(* PLC project DsmEasyConfig *)
(* stored: creationDateTime 2022-10-05T09:23:09.683, modificationDateTime 2022-10-05T09:23:09.683 *)

TYPE DFC_rbr_outA01OL : STRUCT
  DTC : UDINT := 16#140100;
  DFCid : UINT := 471;
  debounceMethod : USINT := TIME_UP_DOWN;
END_STRUCT;
END_TYPE

TYPE DFC_rbr_outA01OT : STRUCT
  DTC : UDINT := 16#140200;
  DFCid : UINT := 472;
  debounceMethod : USINT := TIME_UP_DOWN;
END_STRUCT;
END_TYPE

TYPE DFC_rbr_outA01SCB : STRUCT
  DTC : UDINT := 16#140300;
  DFCid : UINT := 473;
  debounceMethod : USINT := TIME_UP_DOWN;
END_STRUCT;
END_TYPE

TYPE DFC_rbr_outA02OC : STRUCT
  DTC : UDINT := 16#140500;
  DFCid : UINT := 971;
  debounceMethod : USINT := NO_DEBOUNCE;
END_STRUCT;
END_TYPE

TYPE DFC_rbr_outA01SCG : STRUCT
  DTC : UDINT := 16#140400;
  DFCid : UINT := 474;
  debounceMethod : USINT := TIME_UP_DOWN;
END_STRUCT;
END_TYPE

TYPE DFC_rbr_outA02OL : STRUCT
  DTC : UDINT := 16#140600;
  DFCid : UINT := 475;
  debounceMethod : USINT := TIME_UP_DOWN;
END_STRUCT;
END_TYPE

TYPE DFC_rbr_outA02OR : STRUCT
  DTC : UDINT := 16#140700;
  DFCid : UINT := 476;
  debounceMethod : USINT := TIME_UP_DOWN;
END_STRUCT;
END_TYPE

TYPE DFC_rbr_outA02OT : STRUCT
  DTC : UDINT := 16#140800;
  DFCid : UINT := 477;
  debounceMethod : USINT := TIME_UP_DOWN;
END_STRUCT;
END_TYPE

TYPE DFC_rbr_outA02SCB : STRUCT
  DTC : UDINT := 16#140900;
  DFCid : UINT := 478;
  debounceMethod : USINT := TIME_UP_DOWN;
END_STRUCT;
END_TYPE

TYPE DFC_rbr_outA02SCG : STRUCT
  DTC : UDINT := 16#140A00;
  DFCid : UINT := 479;
  debounceMethod : USINT := TIME_UP_DOWN;
END_STRUCT;
END_TYPE

TYPE DFC_rbr_outA03OC : STRUCT
  DTC : UDINT := 16#140B00;
  DFCid : UINT := 973;
  debounceMethod : USINT := NO_DEBOUNCE;
END_STRUCT;
END_TYPE

TYPE DFC_rbr_outA03OL : STRUCT
  DTC : UDINT := 16#140C00;
  DFCid : UINT := 480;
  debounceMethod : USINT := TIME_UP_DOWN;
END_STRUCT;
END_TYPE

TYPE DFC_rbr_outA03OT : STRUCT
  DTC : UDINT := 16#140D00;
  DFCid : UINT := 481;
  debounceMethod : USINT := TIME_UP_DOWN;
END_STRUCT;
END_TYPE

TYPE DFC_rbr_outA03SCB : STRUCT
  DTC : UDINT := 16#140E00;
  DFCid : UINT := 482;
  debounceMethod : USINT := TIME_UP_DOWN;
END_STRUCT;
END_TYPE

TYPE DFC_rbr_outA03SCG : STRUCT
  DTC : UDINT := 16#140F00;
  DFCid : UINT := 483;
  debounceMethod : USINT := TIME_UP_DOWN;
END_STRUCT;
END_TYPE

TYPE DFC_rbr_outA04OC : STRUCT
  DTC : UDINT := 16#141000;
  DFCid : UINT := 975;
  debounceMethod : USINT := NO_DEBOUNCE;
END_STRUCT;
END_TYPE

TYPE DFC_rbr_outA04OL : STRUCT
  DTC : UDINT := 16#141100;
  DFCid : UINT := 484;
  debounceMethod : USINT := TIME_UP_DOWN;
END_STRUCT;
END_TYPE

TYPE DFC_rbr_outA04OT : STRUCT
  DTC : UDINT := 16#141200;
  DFCid : UINT := 485;
  debounceMethod : USINT := TIME_UP_DOWN;
END_STRUCT;
END_TYPE

TYPE DFC_rbr_outA04SCB : STRUCT
  DTC : UDINT := 16#141300;
  DFCid : UINT := 486;
  debounceMethod : USINT := TIME_UP_DOWN;
END_STRUCT;
END_TYPE

TYPE DFC_rbr_outA04SCG : STRUCT
  DTC : UDINT := 16#141400;
  DFCid : UINT := 487;
  debounceMethod : USINT := TIME_UP_DOWN;
END_STRUCT;
END_TYPE

TYPE DFC_rbr_outA05OC : STRUCT
  DTC : UDINT := 16#141500;
  DFCid : UINT := 977;
  debounceMethod : USINT := NO_DEBOUNCE;
END_STRUCT;
END_TYPE

TYPE DFC_rbr_outA05OL : STRUCT
  DTC : UDINT := 16#141600;
  DFCid : UINT := 488;
  debounceMethod : USINT := TIME_UP_DOWN;
END_STRUCT;
END_TYPE

TYPE DFC_rbr_outA05OR : STRUCT
  DTC : UDINT := 16#141700;
  DFCid : UINT := 489;
  debounceMethod : USINT := TIME_UP_DOWN;
END_STRUCT;
END_TYPE

TYPE DFC_rbr_outA05OT : STRUCT
  DTC : UDINT := 16#141800;
  DFCid : UINT := 490;
  debounceMethod : USINT := TIME_UP_DOWN;
END_STRUCT;
END_TYPE

TYPE DFC_rbr_outA05SCB : STRUCT
  DTC : UDINT := 16#141900;
  DFCid : UINT := 491;
  debounceMethod : USINT := TIME_UP_DOWN;
END_STRUCT;
END_TYPE

TYPE DFC_rbr_outA05SCG : STRUCT
  DTC : UDINT := 16#141A00;
  DFCid : UINT := 492;
  debounceMethod : USINT := TIME_UP_DOWN;
END_STRUCT;
END_TYPE

TYPE DFC_rbr_outA06OR : STRUCT
  DTC : UDINT := 16#141C00;
  DFCid : UINT := 494;
  debounceMethod : USINT := TIME_UP_DOWN;
END_STRUCT;
END_TYPE

TYPE DFC_rbr_outA06OT : STRUCT
  DTC : UDINT := 16#141D00;
  DFCid : UINT := 495;
  debounceMethod : USINT := TIME_UP_DOWN;
END_STRUCT;
END_TYPE

TYPE DFC_rbr_outA06SCB : STRUCT
  DTC : UDINT := 16#141E00;
  DFCid : UINT := 496;
  debounceMethod : USINT := TIME_UP_DOWN;
END_STRUCT;
END_TYPE

TYPE DFC_rbr_outA06SCG : STRUCT
  DTC : UDINT := 16#141F00;
  DFCid : UINT := 497;
  debounceMethod : USINT := TIME_UP_DOWN;
END_STRUCT;
END_TYPE

TYPE DFC_rbr_outA07OC : STRUCT
  DTC : UDINT := 16#142000;
  DFCid : UINT := 979;
  debounceMethod : USINT := NO_DEBOUNCE;
END_STRUCT;
END_TYPE

TYPE DFC_rbr_outA07OL : STRUCT
  DTC : UDINT := 16#142100;
  DFCid : UINT := 498;
  debounceMethod : USINT := TIME_UP_DOWN;
END_STRUCT;
END_TYPE

TYPE DFC_rbr_outA07OT : STRUCT
  DTC : UDINT := 16#142200;
  DFCid : UINT := 499;
  debounceMethod : USINT := TIME_UP_DOWN;
END_STRUCT;
END_TYPE

TYPE DFC_rbr_outA07SCB : STRUCT
  DTC : UDINT := 16#142300;
  DFCid : UINT := 500;
  debounceMethod : USINT := TIME_UP_DOWN;
END_STRUCT;
END_TYPE

TYPE DFC_rbr_outA07SCG : STRUCT
  DTC : UDINT := 16#142400;
  DFCid : UINT := 501;
  debounceMethod : USINT := TIME_UP_DOWN;
END_STRUCT;
END_TYPE

TYPE DFC_rbr_outA08OC : STRUCT
  DTC : UDINT := 16#142500;
  DFCid : UINT := 981;
  debounceMethod : USINT := NO_DEBOUNCE;
END_STRUCT;
END_TYPE

TYPE DFC_rbr_outA08OL : STRUCT
  DTC : UDINT := 16#142600;
  DFCid : UINT := 502;
  debounceMethod : USINT := TIME_UP_DOWN;
END_STRUCT;
END_TYPE

TYPE DFC_rbr_outA08OT : STRUCT
  DTC : UDINT := 16#142700;
  DFCid : UINT := 503;
  debounceMethod : USINT := TIME_UP_DOWN;
END_STRUCT;
END_TYPE

TYPE DFC_rbr_outA08SCB : STRUCT
  DTC : UDINT := 16#142800;
  DFCid : UINT := 504;
  debounceMethod : USINT := TIME_UP_DOWN;
END_STRUCT;
END_TYPE

TYPE DFC_rbr_outA08SCG : STRUCT
  DTC : UDINT := 16#142900;
  DFCid : UINT := 505;
  debounceMethod : USINT := TIME_UP_DOWN;
END_STRUCT;
END_TYPE

TYPE DFC_rbr_outA09OC : STRUCT
  DTC : UDINT := 16#142A00;
  DFCid : UINT := 983;
  debounceMethod : USINT := NO_DEBOUNCE;
END_STRUCT;
END_TYPE

TYPE DFC_rbr_outA09OL : STRUCT
  DTC : UDINT := 16#142B00;
  DFCid : UINT := 506;
  debounceMethod : USINT := TIME_UP_DOWN;
END_STRUCT;
END_TYPE

TYPE DFC_rbr_outA09OR : STRUCT
  DTC : UDINT := 16#142C00;
  DFCid : UINT := 507;
  debounceMethod : USINT := TIME_UP_DOWN;
END_STRUCT;
END_TYPE

TYPE DFC_rbr_outA09OT : STRUCT
  DTC : UDINT := 16#142D00;
  DFCid : UINT := 508;
  debounceMethod : USINT := TIME_UP_DOWN;
END_STRUCT;
END_TYPE

TYPE DFC_rbr_outA09SCB : STRUCT
  DTC : UDINT := 16#142E00;
  DFCid : UINT := 509;
  debounceMethod : USINT := TIME_UP_DOWN;
END_STRUCT;
END_TYPE

TYPE DFC_rbr_outA09SCG : STRUCT
  DTC : UDINT := 16#142F00;
  DFCid : UINT := 510;
  debounceMethod : USINT := TIME_UP_DOWN;
END_STRUCT;
END_TYPE

TYPE DFC_rbr_outA10OC : STRUCT
  DTC : UDINT := 16#143000;
  DFCid : UINT := 985;
  debounceMethod : USINT := NO_DEBOUNCE;
END_STRUCT;
END_TYPE

TYPE DFC_rbr_outA10OL : STRUCT
  DTC : UDINT := 16#143100;
  DFCid : UINT := 511;
  debounceMethod : USINT := TIME_UP_DOWN;
END_STRUCT;
END_TYPE

TYPE DFC_rbr_outA10OT : STRUCT
  DTC : UDINT := 16#143200;
  DFCid : UINT := 512;
  debounceMethod : USINT := TIME_UP_DOWN;
END_STRUCT;
END_TYPE

TYPE DFC_rbr_outA10SCB : STRUCT
  DTC : UDINT := 16#143300;
  DFCid : UINT := 513;
  debounceMethod : USINT := TIME_UP_DOWN;
END_STRUCT;
END_TYPE

TYPE DFC_rbr_outA10SCG : STRUCT
  DTC : UDINT := 16#143400;
  DFCid : UINT := 514;
  debounceMethod : USINT := TIME_UP_DOWN;
END_STRUCT;
END_TYPE

TYPE DFC_rbr_outA11OL : STRUCT
  DTC : UDINT := 16#143500;
  DFCid : UINT := 515;
  debounceMethod : USINT := TIME_UP_DOWN;
END_STRUCT;
END_TYPE

TYPE DFC_rbr_outA11OT : STRUCT
  DTC : UDINT := 16#143600;
  DFCid : UINT := 516;
  debounceMethod : USINT := TIME_UP_DOWN;
END_STRUCT;
END_TYPE

TYPE DFC_rbr_outA11SCB : STRUCT
  DTC : UDINT := 16#143700;
  DFCid : UINT := 517;
  debounceMethod : USINT := TIME_UP_DOWN;
END_STRUCT;
END_TYPE

TYPE DFC_rbr_outA11SCG : STRUCT
  DTC : UDINT := 16#143800;
  DFCid : UINT := 518;
  debounceMethod : USINT := TIME_UP_DOWN;
END_STRUCT;
END_TYPE

TYPE DFC_rbr_outA12OR : STRUCT
  DTC : UDINT := 16#143900;
  DFCid : UINT := 519;
  debounceMethod : USINT := TIME_UP_DOWN;
END_STRUCT;
END_TYPE

TYPE DFC_rbr_outA17OC : STRUCT
  DTC : UDINT := 16#144000;
  DFCid : UINT := 987;
  debounceMethod : USINT := NO_DEBOUNCE;
END_STRUCT;
END_TYPE

TYPE DFC_rbr_outA17OL : STRUCT
  DTC : UDINT := 16#144100;
  DFCid : UINT := 526;
  debounceMethod : USINT := TIME_UP_DOWN;
END_STRUCT;
END_TYPE

TYPE DFC_rbr_outA17OR : STRUCT
  DTC : UDINT := 16#144200;
  DFCid : UINT := 527;
  debounceMethod : USINT := TIME_UP_DOWN;
END_STRUCT;
END_TYPE

TYPE DFC_rbr_outA17OT : STRUCT
  DTC : UDINT := 16#144300;
  DFCid : UINT := 528;
  debounceMethod : USINT := TIME_UP_DOWN;
END_STRUCT;
END_TYPE

TYPE DFC_rbr_outA17SCB : STRUCT
  DTC : UDINT := 16#144400;
  DFCid : UINT := 529;
  debounceMethod : USINT := TIME_UP_DOWN;
END_STRUCT;
END_TYPE

TYPE DFC_rbr_outA17SCG : STRUCT
  DTC : UDINT := 16#144500;
  DFCid : UINT := 530;
  debounceMethod : USINT := TIME_UP_DOWN;
END_STRUCT;
END_TYPE

TYPE DFC_rbr_outA18OC : STRUCT
  DTC : UDINT := 16#144600;
  DFCid : UINT := 989;
  debounceMethod : USINT := NO_DEBOUNCE;
END_STRUCT;
END_TYPE

TYPE DFC_rbr_outA18OL : STRUCT
  DTC : UDINT := 16#144700;
  DFCid : UINT := 531;
  debounceMethod : USINT := TIME_UP_DOWN;
END_STRUCT;
END_TYPE

TYPE DFC_rbr_outA18OT : STRUCT
  DTC : UDINT := 16#144800;
  DFCid : UINT := 532;
  debounceMethod : USINT := TIME_UP_DOWN;
END_STRUCT;
END_TYPE

TYPE DFC_rbr_outA18SCB : STRUCT
  DTC : UDINT := 16#144900;
  DFCid : UINT := 533;
  debounceMethod : USINT := TIME_UP_DOWN;
END_STRUCT;
END_TYPE

TYPE DFC_rbr_outA18SCG : STRUCT
  DTC : UDINT := 16#144A00;
  DFCid : UINT := 534;
  debounceMethod : USINT := TIME_UP_DOWN;
END_STRUCT;
END_TYPE

TYPE DFC_rbr_outA19OC : STRUCT
  DTC : UDINT := 16#144B00;
  DFCid : UINT := 991;
  debounceMethod : USINT := NO_DEBOUNCE;
END_STRUCT;
END_TYPE

TYPE DFC_rbr_outA19OL : STRUCT
  DTC : UDINT := 16#144C00;
  DFCid : UINT := 535;
  debounceMethod : USINT := TIME_UP_DOWN;
END_STRUCT;
END_TYPE

TYPE DFC_rbr_outA19OR : STRUCT
  DTC : UDINT := 16#144D00;
  DFCid : UINT := 536;
  debounceMethod : USINT := TIME_UP_DOWN;
END_STRUCT;
END_TYPE

TYPE DFC_rbr_outA19OT : STRUCT
  DTC : UDINT := 16#144E00;
  DFCid : UINT := 537;
  debounceMethod : USINT := TIME_UP_DOWN;
END_STRUCT;
END_TYPE

TYPE DFC_rbr_outA19SCB : STRUCT
  DTC : UDINT := 16#144F00;
  DFCid : UINT := 538;
  debounceMethod : USINT := TIME_UP_DOWN;
END_STRUCT;
END_TYPE

TYPE DFC_rbr_outA19SCG : STRUCT
  DTC : UDINT := 16#145000;
  DFCid : UINT := 539;
  debounceMethod : USINT := TIME_UP_DOWN;
END_STRUCT;
END_TYPE

TYPE DFC_rbr_outA20OC : STRUCT
  DTC : UDINT := 16#145100;
  DFCid : UINT := 993;
  debounceMethod : USINT := NO_DEBOUNCE;
END_STRUCT;
END_TYPE

TYPE DFC_rbr_outA20OL : STRUCT
  DTC : UDINT := 16#145200;
  DFCid : UINT := 540;
  debounceMethod : USINT := TIME_UP_DOWN;
END_STRUCT;
END_TYPE

TYPE DFC_rbr_outA20OR : STRUCT
  DTC : UDINT := 16#145300;
  DFCid : UINT := 541;
  debounceMethod : USINT := TIME_UP_DOWN;
END_STRUCT;
END_TYPE

TYPE DFC_rbr_outA20OT : STRUCT
  DTC : UDINT := 16#145400;
  DFCid : UINT := 542;
  debounceMethod : USINT := TIME_UP_DOWN;
END_STRUCT;
END_TYPE

TYPE DFC_rbr_outA20SCB : STRUCT
  DTC : UDINT := 16#145500;
  DFCid : UINT := 543;
  debounceMethod : USINT := TIME_UP_DOWN;
END_STRUCT;
END_TYPE

TYPE DFC_rbr_outA20SCG : STRUCT
  DTC : UDINT := 16#145600;
  DFCid : UINT := 544;
  debounceMethod : USINT := TIME_UP_DOWN;
END_STRUCT;
END_TYPE

TYPE DFC_rbr_outA31OC : STRUCT
  DTC : UDINT := 16#145700;
  DFCid : UINT := 995;
  debounceMethod : USINT := NO_DEBOUNCE;
END_STRUCT;
END_TYPE

TYPE DFC_rbr_outA31OL : STRUCT
  DTC : UDINT := 16#145800;
  DFCid : UINT := 545;
  debounceMethod : USINT := TIME_UP_DOWN;
END_STRUCT;
END_TYPE

TYPE DFC_rbr_outA31OR : STRUCT
  DTC : UDINT := 16#145900;
  DFCid : UINT := 546;
  debounceMethod : USINT := TIME_UP_DOWN;
END_STRUCT;
END_TYPE

TYPE DFC_rbr_outA31OT : STRUCT
  DTC : UDINT := 16#145A00;
  DFCid : UINT := 547;
  debounceMethod : USINT := TIME_UP_DOWN;
END_STRUCT;
END_TYPE

TYPE DFC_rbr_outA31SCB : STRUCT
  DTC : UDINT := 16#145B00;
  DFCid : UINT := 548;
  debounceMethod : USINT := TIME_UP_DOWN;
END_STRUCT;
END_TYPE

TYPE DFC_rbr_outA31SCG : STRUCT
  DTC : UDINT := 16#145C00;
  DFCid : UINT := 549;
  debounceMethod : USINT := TIME_UP_DOWN;
END_STRUCT;
END_TYPE

TYPE DFC_rbr_outA32OC : STRUCT
  DTC : UDINT := 16#145D00;
  DFCid : UINT := 997;
  debounceMethod : USINT := NO_DEBOUNCE;
END_STRUCT;
END_TYPE

TYPE DFC_rbr_outA32OL : STRUCT
  DTC : UDINT := 16#145E00;
  DFCid : UINT := 550;
  debounceMethod : USINT := TIME_UP_DOWN;
END_STRUCT;
END_TYPE

TYPE DFC_rbr_outA32OR : STRUCT
  DTC : UDINT := 16#145F00;
  DFCid : UINT := 551;
  debounceMethod : USINT := TIME_UP_DOWN;
END_STRUCT;
END_TYPE

TYPE DFC_rbr_outA32OT : STRUCT
  DTC : UDINT := 16#146000;
  DFCid : UINT := 552;
  debounceMethod : USINT := TIME_UP_DOWN;
END_STRUCT;
END_TYPE

TYPE DFC_rbr_outA32SCB : STRUCT
  DTC : UDINT := 16#146100;
  DFCid : UINT := 553;
  debounceMethod : USINT := TIME_UP_DOWN;
END_STRUCT;
END_TYPE

TYPE DFC_rbr_outA32SCG : STRUCT
  DTC : UDINT := 16#146200;
  DFCid : UINT := 554;
  debounceMethod : USINT := TIME_UP_DOWN;
END_STRUCT;
END_TYPE

TYPE DFC_rbr_outA33OC : STRUCT
  DTC : UDINT := 16#146300;
  DFCid : UINT := 999;
  debounceMethod : USINT := NO_DEBOUNCE;
END_STRUCT;
END_TYPE

TYPE DFC_rbr_outA33OL : STRUCT
  DTC : UDINT := 16#146400;
  DFCid : UINT := 555;
  debounceMethod : USINT := TIME_UP_DOWN;
END_STRUCT;
END_TYPE

TYPE DFC_rbr_outA33OR : STRUCT
  DTC : UDINT := 16#146500;
  DFCid : UINT := 556;
  debounceMethod : USINT := TIME_UP_DOWN;
END_STRUCT;
END_TYPE

TYPE DFC_rbr_outA33OT : STRUCT
  DTC : UDINT := 16#146600;
  DFCid : UINT := 557;
  debounceMethod : USINT := TIME_UP_DOWN;
END_STRUCT;
END_TYPE

TYPE DFC_rbr_outA33SCB : STRUCT
  DTC : UDINT := 16#146700;
  DFCid : UINT := 558;
  debounceMethod : USINT := TIME_UP_DOWN;
END_STRUCT;
END_TYPE

TYPE DFC_rbr_outA33SCG : STRUCT
  DTC : UDINT := 16#146800;
  DFCid : UINT := 559;
  debounceMethod : USINT := TIME_UP_DOWN;
END_STRUCT;
END_TYPE

TYPE DFC_rbr_outA34OC : STRUCT
  DTC : UDINT := 16#146900;
  DFCid : UINT := 1001;
  debounceMethod : USINT := NO_DEBOUNCE;
END_STRUCT;
END_TYPE

TYPE DFC_rbr_outA34OL : STRUCT
  DTC : UDINT := 16#146A00;
  DFCid : UINT := 560;
  debounceMethod : USINT := TIME_UP_DOWN;
END_STRUCT;
END_TYPE

TYPE DFC_rbr_outA34OR : STRUCT
  DTC : UDINT := 16#146B00;
  DFCid : UINT := 561;
  debounceMethod : USINT := TIME_UP_DOWN;
END_STRUCT;
END_TYPE

TYPE DFC_rbr_outA34OT : STRUCT
  DTC : UDINT := 16#146C00;
  DFCid : UINT := 562;
  debounceMethod : USINT := TIME_UP_DOWN;
END_STRUCT;
END_TYPE

TYPE DFC_rbr_outA34SCB : STRUCT
  DTC : UDINT := 16#146D00;
  DFCid : UINT := 563;
  debounceMethod : USINT := TIME_UP_DOWN;
END_STRUCT;
END_TYPE

TYPE DFC_rbr_outA34SCG : STRUCT
  DTC : UDINT := 16#146E00;
  DFCid : UINT := 564;
  debounceMethod : USINT := TIME_UP_DOWN;
END_STRUCT;
END_TYPE

TYPE DFC_rbr_outA35OC : STRUCT
  DTC : UDINT := 16#146F00;
  DFCid : UINT := 1003;
  debounceMethod : USINT := NO_DEBOUNCE;
END_STRUCT;
END_TYPE

TYPE DFC_rbr_outA35OL : STRUCT
  DTC : UDINT := 16#147000;
  DFCid : UINT := 565;
  debounceMethod : USINT := TIME_UP_DOWN;
END_STRUCT;
END_TYPE

TYPE DFC_rbr_outA35OR : STRUCT
  DTC : UDINT := 16#147100;
  DFCid : UINT := 566;
  debounceMethod : USINT := TIME_UP_DOWN;
END_STRUCT;
END_TYPE

TYPE DFC_rbr_outA35OT : STRUCT
  DTC : UDINT := 16#147200;
  DFCid : UINT := 567;
  debounceMethod : USINT := TIME_UP_DOWN;
END_STRUCT;
END_TYPE

TYPE DFC_rbr_outA35SCB : STRUCT
  DTC : UDINT := 16#147300;
  DFCid : UINT := 568;
  debounceMethod : USINT := TIME_UP_DOWN;
END_STRUCT;
END_TYPE

TYPE DFC_rbr_outA35SCG : STRUCT
  DTC : UDINT := 16#147400;
  DFCid : UINT := 569;
  debounceMethod : USINT := TIME_UP_DOWN;
END_STRUCT;
END_TYPE

TYPE DFC_rbr_outA46OC : STRUCT
  DTC : UDINT := 16#147500;
  DFCid : UINT := 1005;
  debounceMethod : USINT := NO_DEBOUNCE;
END_STRUCT;
END_TYPE

TYPE DFC_rbr_outA46OL : STRUCT
  DTC : UDINT := 16#147600;
  DFCid : UINT := 570;
  debounceMethod : USINT := TIME_UP_DOWN;
END_STRUCT;
END_TYPE

TYPE DFC_rbr_outA46OR : STRUCT
  DTC : UDINT := 16#147700;
  DFCid : UINT := 571;
  debounceMethod : USINT := TIME_UP_DOWN;
END_STRUCT;
END_TYPE

TYPE DFC_rbr_outA46OT : STRUCT
  DTC : UDINT := 16#147800;
  DFCid : UINT := 572;
  debounceMethod : USINT := TIME_UP_DOWN;
END_STRUCT;
END_TYPE

TYPE DFC_rbr_outA46SCB : STRUCT
  DTC : UDINT := 16#147900;
  DFCid : UINT := 573;
  debounceMethod : USINT := TIME_UP_DOWN;
END_STRUCT;
END_TYPE

TYPE DFC_rbr_outA46SCG : STRUCT
  DTC : UDINT := 16#147A00;
  DFCid : UINT := 574;
  debounceMethod : USINT := TIME_UP_DOWN;
END_STRUCT;
END_TYPE

TYPE DFC_rbr_outA47OC : STRUCT
  DTC : UDINT := 16#147B00;
  DFCid : UINT := 1007;
  debounceMethod : USINT := NO_DEBOUNCE;
END_STRUCT;
END_TYPE

TYPE DFC_rbr_outA47OL : STRUCT
  DTC : UDINT := 16#147C00;
  DFCid : UINT := 575;
  debounceMethod : USINT := TIME_UP_DOWN;
END_STRUCT;
END_TYPE

TYPE DFC_rbr_outA47OR : STRUCT
  DTC : UDINT := 16#147D00;
  DFCid : UINT := 576;
  debounceMethod : USINT := TIME_UP_DOWN;
END_STRUCT;
END_TYPE

TYPE DFC_rbr_outA47OT : STRUCT
  DTC : UDINT := 16#147E00;
  DFCid : UINT := 577;
  debounceMethod : USINT := TIME_UP_DOWN;
END_STRUCT;
END_TYPE

TYPE DFC_rbr_outA47SCB : STRUCT
  DTC : UDINT := 16#147F00;
  DFCid : UINT := 578;
  debounceMethod : USINT := TIME_UP_DOWN;
END_STRUCT;
END_TYPE

TYPE DFC_rbr_outA47SCG : STRUCT
  DTC : UDINT := 16#148000;
  DFCid : UINT := 579;
  debounceMethod : USINT := TIME_UP_DOWN;
END_STRUCT;
END_TYPE

TYPE DFC_rbr_outA48OC : STRUCT
  DTC : UDINT := 16#148100;
  DFCid : UINT := 1009;
  debounceMethod : USINT := NO_DEBOUNCE;
END_STRUCT;
END_TYPE

TYPE DFC_rbr_outA48OL : STRUCT
  DTC : UDINT := 16#148200;
  DFCid : UINT := 580;
  debounceMethod : USINT := TIME_UP_DOWN;
END_STRUCT;
END_TYPE

TYPE DFC_rbr_outA48OR : STRUCT
  DTC : UDINT := 16#148300;
  DFCid : UINT := 581;
  debounceMethod : USINT := TIME_UP_DOWN;
END_STRUCT;
END_TYPE

TYPE DFC_rbr_outA48OT : STRUCT
  DTC : UDINT := 16#148400;
  DFCid : UINT := 582;
  debounceMethod : USINT := TIME_UP_DOWN;
END_STRUCT;
END_TYPE

TYPE DFC_rbr_outA48SCB : STRUCT
  DTC : UDINT := 16#148500;
  DFCid : UINT := 583;
  debounceMethod : USINT := TIME_UP_DOWN;
END_STRUCT;
END_TYPE

TYPE DFC_rbr_outA48SCG : STRUCT
  DTC : UDINT := 16#148600;
  DFCid : UINT := 584;
  debounceMethod : USINT := TIME_UP_DOWN;
END_STRUCT;
END_TYPE

TYPE DFC_rbr_outA49OL : STRUCT
  DTC : UDINT := 16#148700;
  DFCid : UINT := 585;
  debounceMethod : USINT := TIME_UP_DOWN;
END_STRUCT;
END_TYPE

TYPE DFC_rbr_outA49OT : STRUCT
  DTC : UDINT := 16#148800;
  DFCid : UINT := 586;
  debounceMethod : USINT := TIME_UP_DOWN;
END_STRUCT;
END_TYPE

TYPE DFC_rbr_outA49SCB : STRUCT
  DTC : UDINT := 16#148900;
  DFCid : UINT := 587;
  debounceMethod : USINT := TIME_UP_DOWN;
END_STRUCT;
END_TYPE

TYPE DFC_rbr_outA49SCG : STRUCT
  DTC : UDINT := 16#148A00;
  DFCid : UINT := 588;
  debounceMethod : USINT := TIME_UP_DOWN;
END_STRUCT;
END_TYPE

TYPE DFC_rbr_outA50OL : STRUCT
  DTC : UDINT := 16#148B00;
  DFCid : UINT := 589;
  debounceMethod : USINT := TIME_UP_DOWN;
END_STRUCT;
END_TYPE

TYPE DFC_rbr_outA50OT : STRUCT
  DTC : UDINT := 16#148C00;
  DFCid : UINT := 590;
  debounceMethod : USINT := TIME_UP_DOWN;
END_STRUCT;
END_TYPE

TYPE DFC_rbr_outA50SCB : STRUCT
  DTC : UDINT := 16#148D00;
  DFCid : UINT := 591;
  debounceMethod : USINT := TIME_UP_DOWN;
END_STRUCT;
END_TYPE

TYPE DFC_rbr_outA50SCG : STRUCT
  DTC : UDINT := 16#148E00;
  DFCid : UINT := 592;
  debounceMethod : USINT := TIME_UP_DOWN;
END_STRUCT;
END_TYPE

TYPE DFC_rbr_outA51OC : STRUCT
  DTC : UDINT := 16#148F00;
  DFCid : UINT := 1011;
  debounceMethod : USINT := NO_DEBOUNCE;
END_STRUCT;
END_TYPE

TYPE DFC_rbr_outA51OL : STRUCT
  DTC : UDINT := 16#149000;
  DFCid : UINT := 593;
  debounceMethod : USINT := TIME_UP_DOWN;
END_STRUCT;
END_TYPE

TYPE DFC_rbr_outA51OR : STRUCT
  DTC : UDINT := 16#149100;
  DFCid : UINT := 594;
  debounceMethod : USINT := TIME_UP_DOWN;
END_STRUCT;
END_TYPE

TYPE DFC_rbr_outA51OT : STRUCT
  DTC : UDINT := 16#149200;
  DFCid : UINT := 595;
  debounceMethod : USINT := TIME_UP_DOWN;
END_STRUCT;
END_TYPE

TYPE DFC_rbr_outA51SCB : STRUCT
  DTC : UDINT := 16#149300;
  DFCid : UINT := 596;
  debounceMethod : USINT := TIME_UP_DOWN;
END_STRUCT;
END_TYPE

TYPE DFC_rbr_outA51SCG : STRUCT
  DTC : UDINT := 16#149400;
  DFCid : UINT := 597;
  debounceMethod : USINT := TIME_UP_DOWN;
END_STRUCT;
END_TYPE

TYPE DFC_rbr_outA52OC : STRUCT
  DTC : UDINT := 16#149500;
  DFCid : UINT := 1013;
  debounceMethod : USINT := NO_DEBOUNCE;
END_STRUCT;
END_TYPE

TYPE DFC_rbr_outA52OL : STRUCT
  DTC : UDINT := 16#149600;
  DFCid : UINT := 598;
  debounceMethod : USINT := TIME_UP_DOWN;
END_STRUCT;
END_TYPE

TYPE DFC_rbr_outA52OR : STRUCT
  DTC : UDINT := 16#149700;
  DFCid : UINT := 599;
  debounceMethod : USINT := TIME_UP_DOWN;
END_STRUCT;
END_TYPE

TYPE DFC_rbr_outA52OT : STRUCT
  DTC : UDINT := 16#149800;
  DFCid : UINT := 600;
  debounceMethod : USINT := TIME_UP_DOWN;
END_STRUCT;
END_TYPE

TYPE DFC_rbr_outA52SCB : STRUCT
  DTC : UDINT := 16#149900;
  DFCid : UINT := 601;
  debounceMethod : USINT := TIME_UP_DOWN;
END_STRUCT;
END_TYPE

TYPE DFC_rbr_outA52SCG : STRUCT
  DTC : UDINT := 16#149A00;
  DFCid : UINT := 602;
  debounceMethod : USINT := TIME_UP_DOWN;
END_STRUCT;
END_TYPE

TYPE DFC_rbr_outA53OC : STRUCT
  DTC : UDINT := 16#149B00;
  DFCid : UINT := 1015;
  debounceMethod : USINT := NO_DEBOUNCE;
END_STRUCT;
END_TYPE

TYPE DFC_rbr_outA53OL : STRUCT
  DTC : UDINT := 16#149C00;
  DFCid : UINT := 603;
  debounceMethod : USINT := TIME_UP_DOWN;
END_STRUCT;
END_TYPE

TYPE DFC_rbr_outA53OR : STRUCT
  DTC : UDINT := 16#149D00;
  DFCid : UINT := 604;
  debounceMethod : USINT := TIME_UP_DOWN;
END_STRUCT;
END_TYPE

TYPE DFC_rbr_outA53OT : STRUCT
  DTC : UDINT := 16#149E00;
  DFCid : UINT := 605;
  debounceMethod : USINT := TIME_UP_DOWN;
END_STRUCT;
END_TYPE

TYPE DFC_rbr_outA53SCB : STRUCT
  DTC : UDINT := 16#149F00;
  DFCid : UINT := 606;
  debounceMethod : USINT := TIME_UP_DOWN;
END_STRUCT;
END_TYPE

TYPE DFC_rbr_outA53SCG : STRUCT
  DTC : UDINT := 16#14A000;
  DFCid : UINT := 607;
  debounceMethod : USINT := TIME_UP_DOWN;
END_STRUCT;
END_TYPE

TYPE DFC_rbr_outA54OC : STRUCT
  DTC : UDINT := 16#14A100;
  DFCid : UINT := 1017;
  debounceMethod : USINT := NO_DEBOUNCE;
END_STRUCT;
END_TYPE

TYPE DFC_rbr_outA54OL : STRUCT
  DTC : UDINT := 16#14A200;
  DFCid : UINT := 608;
  debounceMethod : USINT := TIME_UP_DOWN;
END_STRUCT;
END_TYPE

TYPE DFC_rbr_outA54OR : STRUCT
  DTC : UDINT := 16#14A300;
  DFCid : UINT := 609;
  debounceMethod : USINT := TIME_UP_DOWN;
END_STRUCT;
END_TYPE

TYPE DFC_rbr_outA54OT : STRUCT
  DTC : UDINT := 16#14A400;
  DFCid : UINT := 610;
  debounceMethod : USINT := TIME_UP_DOWN;
END_STRUCT;
END_TYPE

TYPE DFC_rbr_outA54SCB : STRUCT
  DTC : UDINT := 16#14A500;
  DFCid : UINT := 611;
  debounceMethod : USINT := TIME_UP_DOWN;
END_STRUCT;
END_TYPE

TYPE DFC_rbr_outA54SCG : STRUCT
  DTC : UDINT := 16#14A600;
  DFCid : UINT := 612;
  debounceMethod : USINT := TIME_UP_DOWN;
END_STRUCT;
END_TYPE

TYPE DFC_rbr_outA55OL : STRUCT
  DTC : UDINT := 16#14A700;
  DFCid : UINT := 613;
  debounceMethod : USINT := TIME_UP_DOWN;
END_STRUCT;
END_TYPE

TYPE DFC_rbr_outA55OT : STRUCT
  DTC : UDINT := 16#14A800;
  DFCid : UINT := 614;
  debounceMethod : USINT := TIME_UP_DOWN;
END_STRUCT;
END_TYPE

TYPE DFC_rbr_outA55SCB : STRUCT
  DTC : UDINT := 16#14A900;
  DFCid : UINT := 615;
  debounceMethod : USINT := TIME_UP_DOWN;
END_STRUCT;
END_TYPE

TYPE DFC_rbr_outA55SCG : STRUCT
  DTC : UDINT := 16#14AA00;
  DFCid : UINT := 616;
  debounceMethod : USINT := TIME_UP_DOWN;
END_STRUCT;
END_TYPE

TYPE DFC_rbr_outA56OL : STRUCT
  DTC : UDINT := 16#14AB00;
  DFCid : UINT := 617;
  debounceMethod : USINT := TIME_UP_DOWN;
END_STRUCT;
END_TYPE

TYPE DFC_rbr_outA56OT : STRUCT
  DTC : UDINT := 16#14AC00;
  DFCid : UINT := 618;
  debounceMethod : USINT := TIME_UP_DOWN;
END_STRUCT;
END_TYPE

TYPE DFC_rbr_outA56SCB : STRUCT
  DTC : UDINT := 16#14AD00;
  DFCid : UINT := 619;
  debounceMethod : USINT := TIME_UP_DOWN;
END_STRUCT;
END_TYPE

TYPE DFC_rbr_outA56SCG : STRUCT
  DTC : UDINT := 16#14AE00;
  DFCid : UINT := 620;
  debounceMethod : USINT := TIME_UP_DOWN;
END_STRUCT;
END_TYPE

TYPE DFC_rbr_outA58OL : STRUCT
  DTC : UDINT := 16#14AF00;
  DFCid : UINT := 621;
  debounceMethod : USINT := TIME_UP_DOWN;
END_STRUCT;
END_TYPE

TYPE DFC_rbr_outA58OT : STRUCT
  DTC : UDINT := 16#14B000;
  DFCid : UINT := 622;
  debounceMethod : USINT := TIME_UP_DOWN;
END_STRUCT;
END_TYPE

TYPE DFC_rbr_outA58SCB : STRUCT
  DTC : UDINT := 16#14B100;
  DFCid : UINT := 623;
  debounceMethod : USINT := TIME_UP_DOWN;
END_STRUCT;
END_TYPE

TYPE DFC_rbr_outA58SCG : STRUCT
  DTC : UDINT := 16#14B200;
  DFCid : UINT := 624;
  debounceMethod : USINT := TIME_UP_DOWN;
END_STRUCT;
END_TYPE

TYPE DFC_rbr_outK14OR : STRUCT
  DTC : UDINT := 16#046300;
  DFCid : UINT := 649;
  debounceMethod : USINT := TIME_UP_DOWN;
END_STRUCT;
END_TYPE

TYPE DFC_rbr_outK15OR : STRUCT
  DTC : UDINT := 16#046400;
  DFCid : UINT := 654;
  debounceMethod : USINT := TIME_UP_DOWN;
END_STRUCT;
END_TYPE

TYPE DFC_rbr_outK16OR : STRUCT
  DTC : UDINT := 16#046500;
  DFCid : UINT := 659;
  debounceMethod : USINT := TIME_UP_DOWN;
END_STRUCT;
END_TYPE

TYPE DFC_rbr_outK17OC : STRUCT
  DTC : UDINT := 16#046600;
  DFCid : UINT := 1047;
  debounceMethod : USINT := NO_DEBOUNCE;
END_STRUCT;
END_TYPE

TYPE DFC_rbr_outK17OL : STRUCT
  DTC : UDINT := 16#046700;
  DFCid : UINT := 663;
  debounceMethod : USINT := TIME_UP_DOWN;
END_STRUCT;
END_TYPE

TYPE DFC_rbr_outK17OR : STRUCT
  DTC : UDINT := 16#046800;
  DFCid : UINT := 664;
  debounceMethod : USINT := TIME_UP_DOWN;
END_STRUCT;
END_TYPE

TYPE DFC_rbr_outK17OT : STRUCT
  DTC : UDINT := 16#046900;
  DFCid : UINT := 665;
  debounceMethod : USINT := TIME_UP_DOWN;
END_STRUCT;
END_TYPE

TYPE DFC_rbr_outK17SCB : STRUCT
  DTC : UDINT := 16#046A00;
  DFCid : UINT := 666;
  debounceMethod : USINT := TIME_UP_DOWN;
END_STRUCT;
END_TYPE

TYPE DFC_rbr_outA06OL : STRUCT
  DTC : UDINT := 16#141B00;
  DFCid : UINT := 493;
  debounceMethod : USINT := TIME_UP_DOWN;
END_STRUCT;
END_TYPE

TYPE DFC_rbr_outA16SCB : STRUCT
  DTC : UDINT := 16#143E00;
  DFCid : UINT := 524;
  debounceMethod : USINT := TIME_UP_DOWN;
END_STRUCT;
END_TYPE

TYPE DFC_rbr_outA16SCG : STRUCT
  DTC : UDINT := 16#143F00;
  DFCid : UINT := 525;
  debounceMethod : USINT := TIME_UP_DOWN;
END_STRUCT;
END_TYPE

TYPE DFC_rbr_outA16OL : STRUCT
  DTC : UDINT := 16#143C00;
  DFCid : UINT := 522;
  debounceMethod : USINT := TIME_UP_DOWN;
END_STRUCT;
END_TYPE

TYPE DFC_rbr_outA16OT : STRUCT
  DTC : UDINT := 16#143D00;
  DFCid : UINT := 523;
  debounceMethod : USINT := TIME_UP_DOWN;
END_STRUCT;
END_TYPE

TYPE DFC_rbr_outA12SCB : STRUCT
  DTC : UDINT := 16#143A00;
  DFCid : UINT := 520;
  debounceMethod : USINT := TIME_UP_DOWN;
END_STRUCT;
END_TYPE

TYPE DFC_rbr_outA12SCG : STRUCT
  DTC : UDINT := 16#143B00;
  DFCid : UINT := 521;
  debounceMethod : USINT := TIME_UP_DOWN;
END_STRUCT;
END_TYPE

TYPE DFC_rbr_outK17SCG : STRUCT
  DTC : UDINT := 16#046B00;
  DFCid : UINT := 667;
  debounceMethod : USINT := TIME_UP_DOWN;
END_STRUCT;
END_TYPE

TYPE DFC_rbr_isobusGetStatusParam : STRUCT
  DTC : UDINT := 16#050500;
  DFCid : UINT := 920;
  debounceMethod : USINT := NO_DEBOUNCE;
END_STRUCT;
END_TYPE

TYPE DFC_rbr_isobusRegisterErrClrCallbackParam : STRUCT
  DTC : UDINT := 16#050D00;
  DFCid : UINT := 934;
  debounceMethod : USINT := NO_DEBOUNCE;
END_STRUCT;
END_TYPE

TYPE DFC_rbr_isobusSetCaInfoParam : STRUCT
  DTC : UDINT := 16#051D00;
  DFCid : UINT := 944;
  debounceMethod : USINT := NO_DEBOUNCE;
END_STRUCT;
END_TYPE

TYPE DFC_rbr_isobusRegisterInstancesOverlap : STRUCT
  DTC : UDINT := 16#050E00;
  DFCid : UINT := 935;
  debounceMethod : USINT := NO_DEBOUNCE;
END_STRUCT;
END_TYPE

TYPE DFC_rbr_isobusRegisterInstancesState : STRUCT
  DTC : UDINT := 16#051000;
  DFCid : UINT := 937;
  debounceMethod : USINT := NO_DEBOUNCE;
END_STRUCT;
END_TYPE

TYPE DFC_rbr_isobusRegisterInstancesParam : STRUCT
  DTC : UDINT := 16#050F00;
  DFCid : UINT := 936;
  debounceMethod : USINT := NO_DEBOUNCE;
END_STRUCT;
END_TYPE

TYPE DFC_rbr_isobusSendRequestPGNParam : STRUCT
  DTC : UDINT := 16#051800;
  DFCid : UINT := 939;
  debounceMethod : USINT := NO_DEBOUNCE;
END_STRUCT;
END_TYPE

TYPE DFC_rbr_isobusGetDiagnosticParam : STRUCT
  DTC : UDINT := 16#050300;
  DFCid : UINT := 918;
  debounceMethod : USINT := NO_DEBOUNCE;
END_STRUCT;
END_TYPE

TYPE DFC_rbr_isobusInitDiagnosticParam : STRUCT
  DTC : UDINT := 16#050900;
  DFCid : UINT := 924;
  debounceMethod : USINT := NO_DEBOUNCE;
END_STRUCT;
END_TYPE

TYPE DFC_rbr_isobusInitFailureListParam : STRUCT
  DTC : UDINT := 16#050A00;
  DFCid : UINT := 925;
  debounceMethod : USINT := NO_DEBOUNCE;
END_STRUCT;
END_TYPE

TYPE DFC_rbr_isobusCanRxBufferOverflow : STRUCT
  DTC : UDINT := 16#050100;
  DFCid : UINT := 916;
  debounceMethod : USINT := NO_DEBOUNCE;
END_STRUCT;
END_TYPE

TYPE DFC_rbr_isobusGetRxDataboxStatusParam : STRUCT
  DTC : UDINT := 16#050400;
  DFCid : UINT := 919;
  debounceMethod : USINT := NO_DEBOUNCE;
END_STRUCT;
END_TYPE

TYPE DFC_rbr_isobusSendDataboxParam : STRUCT
  DTC : UDINT := 16#051700;
  DFCid : UINT := 938;
  debounceMethod : USINT := NO_DEBOUNCE;
END_STRUCT;
END_TYPE

TYPE DFC_rbr_isobusInitTxDataboxParam : STRUCT
  DTC : UDINT := 16#050C00;
  DFCid : UINT := 927;
  debounceMethod : USINT := NO_DEBOUNCE;
END_STRUCT;
END_TYPE

TYPE DFC_rbr_isobusRegTxDataboxState : STRUCT
  DTC : UDINT := 16#051600;
  DFCid : UINT := 933;
  debounceMethod : USINT := NO_DEBOUNCE;
END_STRUCT;
END_TYPE

TYPE DFC_rbr_isobusRegTxDataboxParam : STRUCT
  DTC : UDINT := 16#051500;
  DFCid : UINT := 932;
  debounceMethod : USINT := NO_DEBOUNCE;
END_STRUCT;
END_TYPE

TYPE DFC_rbr_isobusRegTxDataboxOverlap : STRUCT
  DTC : UDINT := 16#051400;
  DFCid : UINT := 931;
  debounceMethod : USINT := NO_DEBOUNCE;
END_STRUCT;
END_TYPE

TYPE DFC_rbr_isobusInitRxDataboxParam : STRUCT
  DTC : UDINT := 16#050B00;
  DFCid : UINT := 926;
  debounceMethod : USINT := NO_DEBOUNCE;
END_STRUCT;
END_TYPE

TYPE DFC_rbr_isobusRegRxDataboxState : STRUCT
  DTC : UDINT := 16#051300;
  DFCid : UINT := 930;
  debounceMethod : USINT := NO_DEBOUNCE;
END_STRUCT;
END_TYPE

TYPE DFC_rbr_isobusRegRxDataboxParam : STRUCT
  DTC : UDINT := 16#051200;
  DFCid : UINT := 929;
  debounceMethod : USINT := NO_DEBOUNCE;
END_STRUCT;
END_TYPE

TYPE DFC_rbr_isobusRegRxDataboxOverlap : STRUCT
  DTC : UDINT := 16#051100;
  DFCid : UINT := 928;
  debounceMethod : USINT := NO_DEBOUNCE;
END_STRUCT;
END_TYPE

TYPE DFC_rbr_isobusGetCaAddrParam : STRUCT
  DTC : UDINT := 16#050200;
  DFCid : UINT := 917;
  debounceMethod : USINT := NO_DEBOUNCE;
END_STRUCT;
END_TYPE

TYPE DFC_rbr_isobusSetCaAddrCaUsed : STRUCT
  DTC : UDINT := 16#051900;
  DFCid : UINT := 940;
  debounceMethod : USINT := NO_DEBOUNCE;
END_STRUCT;
END_TYPE

TYPE DFC_rbr_isobusSetCaAddrInvCan : STRUCT
  DTC : UDINT := 16#051B00;
  DFCid : UINT := 942;
  debounceMethod : USINT := NO_DEBOUNCE;
END_STRUCT;
END_TYPE

TYPE DFC_rbr_isobusSetCaAddrParam : STRUCT
  DTC : UDINT := 16#051C00;
  DFCid : UINT := 943;
  debounceMethod : USINT := NO_DEBOUNCE;
END_STRUCT;
END_TYPE

TYPE DFC_rbr_isobusSetCaAddrComm : STRUCT
  DTC : UDINT := 16#051A00;
  DFCid : UINT := 941;
  debounceMethod : USINT := NO_DEBOUNCE;
END_STRUCT;
END_TYPE

TYPE DFC_rbr_isobusSetCaNameParam : STRUCT
  DTC : UDINT := 16#051E00;
  DFCid : UINT := 945;
  debounceMethod : USINT := NO_DEBOUNCE;
END_STRUCT;
END_TYPE

TYPE DFC_rbr_isobusInitCommCaMissing : STRUCT
  DTC : UDINT := 16#050600;
  DFCid : UINT := 921;
  debounceMethod : USINT := NO_DEBOUNCE;
END_STRUCT;
END_TYPE

TYPE DFC_rbr_isobusInitCommState : STRUCT
  DTC : UDINT := 16#050800;
  DFCid : UINT := 923;
  debounceMethod : USINT := NO_DEBOUNCE;
END_STRUCT;
END_TYPE

TYPE DFC_rbr_isobusInitCommParam : STRUCT
  DTC : UDINT := 16#050700;
  DFCid : UINT := 922;
  debounceMethod : USINT := NO_DEBOUNCE;
END_STRUCT;
END_TYPE

TYPE DFC_rbr_mo_OV_VSS1 : STRUCT
  DTC : UDINT := 16#080100;
  DFCid : UINT := 1156;
  debounceMethod : USINT := NO_DEBOUNCE;
END_STRUCT;
END_TYPE

TYPE DFC_rbr_mo_UV_VSS1 : STRUCT
  DTC : UDINT := 16#080200;
  DFCid : UINT := 1158;
  debounceMethod : USINT := NO_DEBOUNCE;
END_STRUCT;
END_TYPE

TYPE DFC_rbr_mo_OV_VSS2 : STRUCT
  DTC : UDINT := 16#080300;
  DFCid : UINT := 1157;
  debounceMethod : USINT := NO_DEBOUNCE;
END_STRUCT;
END_TYPE

TYPE DFC_rbr_mo_UV_VSS2 : STRUCT
  DTC : UDINT := 16#080400;
  DFCid : UINT := 1159;
  debounceMethod : USINT := NO_DEBOUNCE;
END_STRUCT;
END_TYPE

TYPE DFC_rbr_mo_OV_VSS3 : STRUCT
  DTC : UDINT := 16#080500;
  DFCid : UINT := 458;
  debounceMethod : USINT := TIME_UP_DOWN;
END_STRUCT;
END_TYPE

TYPE DFC_rbr_mo_UV_VSS3 : STRUCT
  DTC : UDINT := 16#080600;
  DFCid : UINT := 469;
  debounceMethod : USINT := TIME_UP_DOWN;
END_STRUCT;
END_TYPE

TYPE DFC_rbr_mo_OV_VSS4 : STRUCT
  DTC : UDINT := 16#080700;
  DFCid : UINT := 459;
  debounceMethod : USINT := TIME_UP_DOWN;
END_STRUCT;
END_TYPE

TYPE DFC_rbr_mo_UV_VSS4 : STRUCT
  DTC : UDINT := 16#080800;
  DFCid : UINT := 470;
  debounceMethod : USINT := TIME_UP_DOWN;
END_STRUCT;
END_TYPE

TYPE DFC_rbr_mo_OV_UBAT_MON : STRUCT
  DTC : UDINT := 16#080900;
  DFCid : UINT := 451;
  debounceMethod : USINT := TIME_UP_DOWN;
END_STRUCT;
END_TYPE

TYPE DFC_rbr_mo_OV_UBRM24_MON : STRUCT
  DTC : UDINT := 16#080A00;
  DFCid : UINT := 454;
  debounceMethod : USINT := TIME_UP_DOWN;
END_STRUCT;
END_TYPE

TYPE DFC_rbr_mo_OV_UBRM24_LOADS : STRUCT
  DTC : UDINT := 16#080C00;
  DFCid : UINT := 453;
  debounceMethod : USINT := TIME_UP_DOWN;
END_STRUCT;
END_TYPE

TYPE DFC_rbr_mo_DvUBAT_FWs : STRUCT
  DTC : UDINT := 16#080D00;
  DFCid : UINT := 446;
  debounceMethod : USINT := TIME_UP_DOWN;
END_STRUCT;
END_TYPE

TYPE DFC_rbr_mo_OVWarn_VPR6 : STRUCT
  DTC : UDINT := 16#081200;
  DFCid : UINT := 448;
  debounceMethod : USINT := TIME_UP_DOWN;
END_STRUCT;
END_TYPE

TYPE DFC_rbr_mo_OVErr_VPR6 : STRUCT
  DTC : UDINT := 16#081100;
  DFCid : UINT := 447;
  debounceMethod : USINT := TIME_UP_DOWN;
END_STRUCT;
END_TYPE

TYPE DFC_rbr_mo_OV_VPR6 : STRUCT
  DTC : UDINT := 16#082000;
  DFCid : UINT := 457;
  debounceMethod : USINT := TIME_UP_DOWN;
END_STRUCT;
END_TYPE

TYPE DFC_rbr_mo_UV_VPR6 : STRUCT
  DTC : UDINT := 16#081300;
  DFCid : UINT := 468;
  debounceMethod : USINT := TIME_UP_DOWN;
END_STRUCT;
END_TYPE

TYPE DFC_rbr_mo_Temp1_HTWarn : STRUCT
  DTC : UDINT := 16#081600;
  DFCid : UINT := 461;
  debounceMethod : USINT := TIME_UP_DOWN;
END_STRUCT;
END_TYPE

TYPE DFC_rbr_mo_Temp1_HTErr : STRUCT
  DTC : UDINT := 16#081700;
  DFCid : UINT := 460;
  debounceMethod : USINT := TIME_UP_DOWN;
END_STRUCT;
END_TYPE

TYPE DFC_rbr_mo_Temp2_HTWarn : STRUCT
  DTC : UDINT := 16#081800;
  DFCid : UINT := 463;
  debounceMethod : USINT := TIME_UP_DOWN;
END_STRUCT;
END_TYPE

TYPE DFC_rbr_mo_OV_UBRM24_FLEXIN : STRUCT
  DTC : UDINT := 16#082300;
  DFCid : UINT := 452;
  debounceMethod : USINT := TIME_UP_DOWN;
END_STRUCT;
END_TYPE

TYPE DFC_rbr_mo_UV_VDD5 : STRUCT
  DTC : UDINT := 16#082500;
  DFCid : UINT := 466;
  debounceMethod : USINT := TIME_UP_DOWN;
END_STRUCT;
END_TYPE

TYPE DFC_rbr_mo_UV_VDD5_IN : STRUCT
  DTC : UDINT := 16#082700;
  DFCid : UINT := 467;
  debounceMethod : USINT := TIME_UP_DOWN;
END_STRUCT;
END_TYPE

TYPE DFC_rbr_mo_OV_VDD5_IN : STRUCT
  DTC : UDINT := 16#082600;
  DFCid : UINT := 456;
  debounceMethod : USINT := TIME_UP_DOWN;
END_STRUCT;
END_TYPE

TYPE DFC_rbr_mo_OV_VDD5 : STRUCT
  DTC : UDINT := 16#082400;
  DFCid : UINT := 455;
  debounceMethod : USINT := TIME_UP_DOWN;
END_STRUCT;
END_TYPE

TYPE DFC_rbr_mo_OV_SAV_LSS_MEAS_CLUSTER_1_3 : STRUCT
  DTC : UDINT := 16#082A00;
  DFCid : UINT := 449;
  debounceMethod : USINT := TIME_UP_DOWN;
END_STRUCT;
END_TYPE

TYPE DFC_rbr_mo_OV_SAV_LSS_MEAS_CLUSTER_2 : STRUCT
  DTC : UDINT := 16#082800;
  DFCid : UINT := 450;
  debounceMethod : USINT := TIME_UP_DOWN;
END_STRUCT;
END_TYPE

TYPE DFC_rbr_mo_UV_SAV_LSS_MEAS_CLUSTER_2 : STRUCT
  DTC : UDINT := 16#082900;
  DFCid : UINT := 465;
  debounceMethod : USINT := TIME_UP_DOWN;
END_STRUCT;
END_TYPE

TYPE DFC_rbr_moOV_FirstConstADC : STRUCT
  DTC : UDINT := 16#082C00;
  DFCid : UINT := 963;
  debounceMethod : USINT := NO_DEBOUNCE;
END_STRUCT;
END_TYPE

TYPE DFC_rbr_moUV_FirstConstADC : STRUCT
  DTC : UDINT := 16#082D00;
  DFCid : UINT := 965;
  debounceMethod : USINT := NO_DEBOUNCE;
END_STRUCT;
END_TYPE

TYPE DFC_rbr_moOV_SecondConstADC : STRUCT
  DTC : UDINT := 16#082E00;
  DFCid : UINT := 964;
  debounceMethod : USINT := NO_DEBOUNCE;
END_STRUCT;
END_TYPE

TYPE DFC_rbr_moUV_SecondConstADC : STRUCT
  DTC : UDINT := 16#082F00;
  DFCid : UINT := 966;
  debounceMethod : USINT := NO_DEBOUNCE;
END_STRUCT;
END_TYPE

TYPE DFC_rbr_mo_Temp2_HTErr : STRUCT
  DTC : UDINT := 16#081900;
  DFCid : UINT := 462;
  debounceMethod : USINT := TIME_UP_DOWN;
END_STRUCT;
END_TYPE

TYPE DFC_rbr_mo_UV_SAV_LSS_MEAS_CLUSTER_1_3 : STRUCT
  DTC : UDINT := 16#082B00;
  DFCid : UINT := 464;
  debounceMethod : USINT := TIME_UP_DOWN;
END_STRUCT;
END_TYPE

TYPE DFC_rbr_mo_adcPDD_fail : STRUCT
  DTC : UDINT := 16#083000;
  DFCid : UINT := 969;
  debounceMethod : USINT := NO_DEBOUNCE;
END_STRUCT;
END_TYPE

TYPE DFC_rbr_canInitParam : STRUCT
  DTC : UDINT := 16#020800;
  DFCid : UINT := 830;
  debounceMethod : USINT := NO_DEBOUNCE;
END_STRUCT;
END_TYPE

TYPE DFC_rbr_canSendDataParam : STRUCT
  DTC : UDINT := 16#022500;
  DFCid : UINT := 858;
  debounceMethod : USINT := NO_DEBOUNCE;
END_STRUCT;
END_TYPE

TYPE DFC_rbr_canSendDataBufOvfl : STRUCT
  DTC : UDINT := 16#022400;
  DFCid : UINT := 857;
  debounceMethod : USINT := NO_DEBOUNCE;
END_STRUCT;
END_TYPE

TYPE DFC_rbr_canRegTxBufParam : STRUCT
  DTC : UDINT := 16#021C00;
  DFCid : UINT := 851;
  debounceMethod : USINT := NO_DEBOUNCE;
END_STRUCT;
END_TYPE

TYPE DFC_rbr_canRegTxBufInvState : STRUCT
  DTC : UDINT := 16#021A00;
  DFCid : UINT := 849;
  debounceMethod : USINT := NO_DEBOUNCE;
END_STRUCT;
END_TYPE

TYPE DFC_rbr_canRegRxCallbParam : STRUCT
  DTC : UDINT := 16#021500;
  DFCid : UINT := 844;
  debounceMethod : USINT := NO_DEBOUNCE;
END_STRUCT;
END_TYPE

TYPE DFC_rbr_canRegRxCallbInvState : STRUCT
  DTC : UDINT := 16#021400;
  DFCid : UINT := 843;
  debounceMethod : USINT := NO_DEBOUNCE;
END_STRUCT;
END_TYPE

TYPE DFC_rbr_canRegBusOffCallbParam : STRUCT
  DTC : UDINT := 16#021000;
  DFCid : UINT := 839;
  debounceMethod : USINT := NO_DEBOUNCE;
END_STRUCT;
END_TYPE

TYPE DFC_rbr_canRegBusOffCallbInvState : STRUCT
  DTC : UDINT := 16#020F00;
  DFCid : UINT := 838;
  debounceMethod : USINT := NO_DEBOUNCE;
END_STRUCT;
END_TYPE

TYPE DFC_rbr_canRegRxDataboxParam : STRUCT
  DTC : UDINT := 16#021900;
  DFCid : UINT := 848;
  debounceMethod : USINT := NO_DEBOUNCE;
END_STRUCT;
END_TYPE

TYPE DFC_rbr_canRegRxDataboxInvState : STRUCT
  DTC : UDINT := 16#021700;
  DFCid : UINT := 846;
  debounceMethod : USINT := NO_DEBOUNCE;
END_STRUCT;
END_TYPE

TYPE DFC_rbr_canRegRxBufParam : STRUCT
  DTC : UDINT := 16#021300;
  DFCid : UINT := 842;
  debounceMethod : USINT := NO_DEBOUNCE;
END_STRUCT;
END_TYPE

TYPE DFC_rbr_canRegRxBufInvState : STRUCT
  DTC : UDINT := 16#021100;
  DFCid : UINT := 840;
  debounceMethod : USINT := NO_DEBOUNCE;
END_STRUCT;
END_TYPE

TYPE DFC_rbr_canInitRxDataboxParam : STRUCT
  DTC : UDINT := 16#020A00;
  DFCid : UINT := 832;
  debounceMethod : USINT := NO_DEBOUNCE;
END_STRUCT;
END_TYPE

TYPE DFC_rbr_canGetDataParam : STRUCT
  DTC : UDINT := 16#020400;
  DFCid : UINT := 824;
  debounceMethod : USINT := NO_DEBOUNCE;
END_STRUCT;
END_TYPE

TYPE DFC_rbr_canGetDataNoBuf : STRUCT
  DTC : UDINT := 16#020300;
  DFCid : UINT := 823;
  debounceMethod : USINT := NO_DEBOUNCE;
END_STRUCT;
END_TYPE

TYPE DFC_rbr_canGetDataboxParam : STRUCT
  DTC : UDINT := 16#020200;
  DFCid : UINT := 826;
  debounceMethod : USINT := NO_DEBOUNCE;
END_STRUCT;
END_TYPE

TYPE DFC_rbr_canGetDataboxNoInit : STRUCT
  DTC : UDINT := 16#020100;
  DFCid : UINT := 825;
  debounceMethod : USINT := NO_DEBOUNCE;
END_STRUCT;
END_TYPE

TYPE DFC_rbr_canInitTxDataboxParam : STRUCT
  DTC : UDINT := 16#020B00;
  DFCid : UINT := 833;
  debounceMethod : USINT := NO_DEBOUNCE;
END_STRUCT;
END_TYPE

TYPE DFC_rbr_canIsDataboxFreeParam : STRUCT
  DTC : UDINT := 16#020D00;
  DFCid : UINT := 836;
  debounceMethod : USINT := NO_DEBOUNCE;
END_STRUCT;
END_TYPE

TYPE DFC_rbr_canIsDataboxFreeNoInit : STRUCT
  DTC : UDINT := 16#020C00;
  DFCid : UINT := 835;
  debounceMethod : USINT := NO_DEBOUNCE;
END_STRUCT;
END_TYPE

TYPE DFC_rbr_canSendDataboxParam : STRUCT
  DTC : UDINT := 16#022300;
  DFCid : UINT := 860;
  debounceMethod : USINT := NO_DEBOUNCE;
END_STRUCT;
END_TYPE

TYPE DFC_rbr_canSendDataboxNoInit : STRUCT
  DTC : UDINT := 16#022200;
  DFCid : UINT := 859;
  debounceMethod : USINT := NO_DEBOUNCE;
END_STRUCT;
END_TYPE

TYPE DFC_rbr_canRegTxDataboxParam : STRUCT
  DTC : UDINT := 16#022000;
  DFCid : UINT := 855;
  debounceMethod : USINT := NO_DEBOUNCE;
END_STRUCT;
END_TYPE

TYPE DFC_rbr_canRegTxDataboxInvState : STRUCT
  DTC : UDINT := 16#021E00;
  DFCid : UINT := 853;
  debounceMethod : USINT := NO_DEBOUNCE;
END_STRUCT;
END_TYPE

TYPE DFC_rbr_canIsTxEmptyParam : STRUCT
  DTC : UDINT := 16#020E00;
  DFCid : UINT := 837;
  debounceMethod : USINT := NO_DEBOUNCE;
END_STRUCT;
END_TYPE

TYPE DFC_rbr_canRegRxDataboxInvNumb : STRUCT
  DTC : UDINT := 16#021600;
  DFCid : UINT := 845;
  debounceMethod : USINT := NO_DEBOUNCE;
END_STRUCT;
END_TYPE

TYPE DFC_rbr_canRegTxDataboxInvNumb : STRUCT
  DTC : UDINT := 16#021D00;
  DFCid : UINT := 852;
  debounceMethod : USINT := NO_DEBOUNCE;
END_STRUCT;
END_TYPE

TYPE DFC_rbr_canGetStatusParam : STRUCT
  DTC : UDINT := 16#020600;
  DFCid : UINT := 828;
  debounceMethod : USINT := NO_DEBOUNCE;
END_STRUCT;
END_TYPE

TYPE DFC_rbr_canGetTxBufStatusParam : STRUCT
  DTC : UDINT := 16#020700;
  DFCid : UINT := 829;
  debounceMethod : USINT := NO_DEBOUNCE;
END_STRUCT;
END_TYPE

TYPE DFC_rbr_canResetTxBufParam : STRUCT
  DTC : UDINT := 16#022100;
  DFCid : UINT := 856;
  debounceMethod : USINT := NO_DEBOUNCE;
END_STRUCT;
END_TYPE

TYPE DFC_rbr_canStopParam : STRUCT
  DTC : UDINT := 16#022800;
  DFCid : UINT := 863;
  debounceMethod : USINT := NO_DEBOUNCE;
END_STRUCT;
END_TYPE

TYPE DFC_rbr_canStartParam : STRUCT
  DTC : UDINT := 16#022700;
  DFCid : UINT := 862;
  debounceMethod : USINT := NO_DEBOUNCE;
END_STRUCT;
END_TYPE

TYPE DFC_rbr_canRegRxBufOverlap : STRUCT
  DTC : UDINT := 16#021200;
  DFCid : UINT := 841;
  debounceMethod : USINT := NO_DEBOUNCE;
END_STRUCT;
END_TYPE

TYPE DFC_rbr_canRegTxBufOverlap : STRUCT
  DTC : UDINT := 16#021B00;
  DFCid : UINT := 850;
  debounceMethod : USINT := NO_DEBOUNCE;
END_STRUCT;
END_TYPE

TYPE DFC_rbr_canRegTxDataboxOverlap : STRUCT
  DTC : UDINT := 16#021F00;
  DFCid : UINT := 854;
  debounceMethod : USINT := NO_DEBOUNCE;
END_STRUCT;
END_TYPE

TYPE DFC_rbr_canRegRxDataboxOverlap : STRUCT
  DTC : UDINT := 16#021800;
  DFCid : UINT := 847;
  debounceMethod : USINT := NO_DEBOUNCE;
END_STRUCT;
END_TYPE

TYPE DFC_rbr_canInitRxDataboxOverlap : STRUCT
  DTC : UDINT := 16#020900;
  DFCid : UINT := 831;
  debounceMethod : USINT := NO_DEBOUNCE;
END_STRUCT;
END_TYPE

TYPE DFC_rbr_canSetTxCycleParam : STRUCT
  DTC : UDINT := 16#022600;
  DFCid : UINT := 861;
  debounceMethod : USINT := NO_DEBOUNCE;
END_STRUCT;
END_TYPE

TYPE DFC_rbr_dsmNumDTCJ1939 : STRUCT
  DTC : UDINT := 16#071300;
  DFCid : UINT := 876;
  debounceMethod : USINT := NO_DEBOUNCE;
END_STRUCT;
END_TYPE

TYPE DFC_rbr_dsmGetDTCJ1939 : STRUCT
  DTC : UDINT := 16#070300;
  DFCid : UINT := 872;
  debounceMethod : USINT := NO_DEBOUNCE;
END_STRUCT;
END_TYPE

TYPE DFC_rbr_dsmgetDFCStatus : STRUCT
  DTC : UDINT := 16#071100;
  DFCid : UINT := 880;
  debounceMethod : USINT := NO_DEBOUNCE;
END_STRUCT;
END_TYPE

TYPE DFC_rbr_dsmtestErrorDFC : STRUCT
  DTC : UDINT := 16#071200;
  DFCid : UINT := 881;
  debounceMethod : USINT := NO_DEBOUNCE;
END_STRUCT;
END_TYPE

TYPE DFC_rbr_dsmGetErrors : STRUCT
  DTC : UDINT := 16#070100;
  DFCid : UINT := 873;
  debounceMethod : USINT := NO_DEBOUNCE;
END_STRUCT;
END_TYPE

TYPE DFC_rbr_dsmDelDTCJ1939 : STRUCT
  DTC : UDINT := 16#070400;
  DFCid : UINT := 869;
  debounceMethod : USINT := NO_DEBOUNCE;
END_STRUCT;
END_TYPE

TYPE DFC_rbr_dsmGetNumErrors : STRUCT
  DTC : UDINT := 16#070200;
  DFCid : UINT := 874;
  debounceMethod : USINT := NO_DEBOUNCE;
END_STRUCT;
END_TYPE

TYPE DFC_rbr_dsmGetDFES : STRUCT
  DTC : UDINT := 16#070500;
  DFCid : UINT := 871;
  debounceMethod : USINT := NO_DEBOUNCE;
END_STRUCT;
END_TYPE

TYPE DFC_rbr_dsmTesterror : STRUCT
  DTC : UDINT := 16#070600;
  DFCid : UINT := 877;
  debounceMethod : USINT := NO_DEBOUNCE;
END_STRUCT;
END_TYPE

TYPE DFC_rbr_dsmDelErrors : STRUCT
  DTC : UDINT := 16#070700;
  DFCid : UINT := 870;
  debounceMethod : USINT := NO_DEBOUNCE;
END_STRUCT;
END_TYPE

TYPE DFC_rbr_dsmUpdateDebError : STRUCT
  DTC : UDINT := 16#070800;
  DFCid : UINT := 878;
  debounceMethod : USINT := NO_DEBOUNCE;
END_STRUCT;
END_TYPE

TYPE DFC_rbr_dsmUpdateError : STRUCT
  DTC : UDINT := 16#070900;
  DFCid : UINT := 879;
  debounceMethod : USINT := NO_DEBOUNCE;
END_STRUCT;
END_TYPE

TYPE DFC_rbr_memGetStatus : STRUCT
  DTC : UDINT := 16#060300;
  DFCid : UINT := 954;
  debounceMethod : USINT := NO_DEBOUNCE;
END_STRUCT;
END_TYPE

TYPE DFC_rbr_memReadBlock : STRUCT
  DTC : UDINT := 16#060200;
  DFCid : UINT := 958;
  debounceMethod : USINT := NO_DEBOUNCE;
END_STRUCT;
END_TYPE

TYPE DFC_rbr_memWriteBlock : STRUCT
  DTC : UDINT := 16#060100;
  DFCid : UINT := 962;
  debounceMethod : USINT := NO_DEBOUNCE;
END_STRUCT;
END_TYPE

TYPE DFC_rbr_canIpduGroupControl : STRUCT
  DTC : UDINT := 16#022D00;
  DFCid : UINT := 834;
  debounceMethod : USINT := NO_DEBOUNCE;
END_STRUCT;
END_TYPE

TYPE DFC_rbr_can_ClearIpduGroup : STRUCT
  DTC : UDINT := 16#022C00;
  DFCid : UINT := 864;
  debounceMethod : USINT := NO_DEBOUNCE;
END_STRUCT;
END_TYPE

TYPE DFC_rbr_can_SetIpduGroup : STRUCT
  DTC : UDINT := 16#022B00;
  DFCid : UINT := 867;
  debounceMethod : USINT := NO_DEBOUNCE;
END_STRUCT;
END_TYPE

TYPE DFC_rbr_can_ReceiveSignal : STRUCT
  DTC : UDINT := 16#022A00;
  DFCid : UINT := 865;
  debounceMethod : USINT := NO_DEBOUNCE;
END_STRUCT;
END_TYPE

TYPE DFC_rbr_can_SendSignal : STRUCT
  DTC : UDINT := 16#022900;
  DFCid : UINT := 866;
  debounceMethod : USINT := NO_DEBOUNCE;
END_STRUCT;
END_TYPE

TYPE DFC_rbr_canGetRxBufStatusParam : STRUCT
  DTC : UDINT := 16#020500;
  DFCid : UINT := 827;
  debounceMethod : USINT := NO_DEBOUNCE;
END_STRUCT;
END_TYPE

TYPE DFC_rbr_inK65ShuntSCB : STRUCT
  DTC : UDINT := 16#03D700;
  DFCid : UINT := 430;
  debounceMethod : USINT := TIME_UP_DOWN;
END_STRUCT;
END_TYPE

TYPE DFC_rbr_inK65AicSCG : STRUCT
  DTC : UDINT := 16#03D600;
  DFCid : UINT := 426;
  debounceMethod : USINT := TIME_UP_DOWN;
END_STRUCT;
END_TYPE

TYPE DFC_rbr_inK65AicSCB : STRUCT
  DTC : UDINT := 16#03D500;
  DFCid : UINT := 425;
  debounceMethod : USINT := TIME_UP_DOWN;
END_STRUCT;
END_TYPE

TYPE DFC_rbr_inK64ShuntSCB : STRUCT
  DTC : UDINT := 16#03D400;
  DFCid : UINT := 424;
  debounceMethod : USINT := TIME_UP_DOWN;
END_STRUCT;
END_TYPE

TYPE DFC_rbr_inK64AicSCG : STRUCT
  DTC : UDINT := 16#03D300;
  DFCid : UINT := 420;
  debounceMethod : USINT := TIME_UP_DOWN;
END_STRUCT;
END_TYPE

TYPE DFC_rbr_inK64AicSCB : STRUCT
  DTC : UDINT := 16#03D200;
  DFCid : UINT := 419;
  debounceMethod : USINT := TIME_UP_DOWN;
END_STRUCT;
END_TYPE

TYPE DFC_rbr_inK63ShuntSCB : STRUCT
  DTC : UDINT := 16#03D100;
  DFCid : UINT := 418;
  debounceMethod : USINT := TIME_UP_DOWN;
END_STRUCT;
END_TYPE

TYPE DFC_rbr_inK63AicSCG : STRUCT
  DTC : UDINT := 16#03D000;
  DFCid : UINT := 414;
  debounceMethod : USINT := TIME_UP_DOWN;
END_STRUCT;
END_TYPE

TYPE DFC_rbr_inK63AicSCB : STRUCT
  DTC : UDINT := 16#03CF00;
  DFCid : UINT := 413;
  debounceMethod : USINT := TIME_UP_DOWN;
END_STRUCT;
END_TYPE

TYPE DFC_rbr_inK45ShuntSCB : STRUCT
  DTC : UDINT := 16#03CE00;
  DFCid : UINT := 370;
  debounceMethod : USINT := TIME_UP_DOWN;
END_STRUCT;
END_TYPE

TYPE DFC_rbr_inK45AicSCG : STRUCT
  DTC : UDINT := 16#03CD00;
  DFCid : UINT := 366;
  debounceMethod : USINT := TIME_UP_DOWN;
END_STRUCT;
END_TYPE

TYPE DFC_rbr_inK45AicSCB : STRUCT
  DTC : UDINT := 16#03CC00;
  DFCid : UINT := 365;
  debounceMethod : USINT := TIME_UP_DOWN;
END_STRUCT;
END_TYPE

TYPE DFC_rbr_inK44ShuntSCB : STRUCT
  DTC : UDINT := 16#03CB00;
  DFCid : UINT := 364;
  debounceMethod : USINT := TIME_UP_DOWN;
END_STRUCT;
END_TYPE

TYPE DFC_rbr_inK44AicSCG : STRUCT
  DTC : UDINT := 16#03CA00;
  DFCid : UINT := 360;
  debounceMethod : USINT := TIME_UP_DOWN;
END_STRUCT;
END_TYPE

TYPE DFC_rbr_inK44AicSCB : STRUCT
  DTC : UDINT := 16#03C900;
  DFCid : UINT := 359;
  debounceMethod : USINT := TIME_UP_DOWN;
END_STRUCT;
END_TYPE

TYPE DFC_rbr_inK42ShuntSCB : STRUCT
  DTC : UDINT := 16#03C800;
  DFCid : UINT := 355;
  debounceMethod : USINT := TIME_UP_DOWN;
END_STRUCT;
END_TYPE

TYPE DFC_rbr_inK42AicSCG : STRUCT
  DTC : UDINT := 16#03C700;
  DFCid : UINT := 351;
  debounceMethod : USINT := TIME_UP_DOWN;
END_STRUCT;
END_TYPE

TYPE DFC_rbr_inK42AicSCB : STRUCT
  DTC : UDINT := 16#03C600;
  DFCid : UINT := 350;
  debounceMethod : USINT := TIME_UP_DOWN;
END_STRUCT;
END_TYPE

TYPE DFC_rbr_inK41ShuntSCB : STRUCT
  DTC : UDINT := 16#03C500;
  DFCid : UINT := 349;
  debounceMethod : USINT := TIME_UP_DOWN;
END_STRUCT;
END_TYPE

TYPE DFC_rbr_inK41AicSCG : STRUCT
  DTC : UDINT := 16#03C400;
  DFCid : UINT := 345;
  debounceMethod : USINT := TIME_UP_DOWN;
END_STRUCT;
END_TYPE

TYPE DFC_rbr_inK41AicSCB : STRUCT
  DTC : UDINT := 16#03C300;
  DFCid : UINT := 344;
  debounceMethod : USINT := TIME_UP_DOWN;
END_STRUCT;
END_TYPE

TYPE DFC_rbr_inK40ShuntSCB : STRUCT
  DTC : UDINT := 16#03C200;
  DFCid : UINT := 343;
  debounceMethod : USINT := TIME_UP_DOWN;
END_STRUCT;
END_TYPE

TYPE DFC_rbr_inK40AicSCG : STRUCT
  DTC : UDINT := 16#03C100;
  DFCid : UINT := 339;
  debounceMethod : USINT := TIME_UP_DOWN;
END_STRUCT;
END_TYPE

TYPE DFC_rbr_inK40AicSCB : STRUCT
  DTC : UDINT := 16#03C000;
  DFCid : UINT := 338;
  debounceMethod : USINT := TIME_UP_DOWN;
END_STRUCT;
END_TYPE

TYPE DFC_rbr_inK39ShuntSCB : STRUCT
  DTC : UDINT := 16#03BF00;
  DFCid : UINT := 337;
  debounceMethod : USINT := TIME_UP_DOWN;
END_STRUCT;
END_TYPE

TYPE DFC_rbr_inK39AicSCG : STRUCT
  DTC : UDINT := 16#03BE00;
  DFCid : UINT := 333;
  debounceMethod : USINT := TIME_UP_DOWN;
END_STRUCT;
END_TYPE

TYPE DFC_rbr_inK39AicSCB : STRUCT
  DTC : UDINT := 16#03BD00;
  DFCid : UINT := 332;
  debounceMethod : USINT := TIME_UP_DOWN;
END_STRUCT;
END_TYPE

TYPE DFC_rbr_inK38ShuntSCB : STRUCT
  DTC : UDINT := 16#03BC00;
  DFCid : UINT := 331;
  debounceMethod : USINT := TIME_UP_DOWN;
END_STRUCT;
END_TYPE

TYPE DFC_rbr_inK38AicSCG : STRUCT
  DTC : UDINT := 16#03BB00;
  DFCid : UINT := 327;
  debounceMethod : USINT := TIME_UP_DOWN;
END_STRUCT;
END_TYPE

TYPE DFC_rbr_inK38AicSCB : STRUCT
  DTC : UDINT := 16#03BA00;
  DFCid : UINT := 326;
  debounceMethod : USINT := TIME_UP_DOWN;
END_STRUCT;
END_TYPE

TYPE DFC_rbr_inK35SCG : STRUCT
  DTC : UDINT := 16#03B900;
  DFCid : UINT := 316;
  debounceMethod : USINT := TIME_UP_DOWN;
END_STRUCT;
END_TYPE

TYPE DFC_rbr_inK35SCB : STRUCT
  DTC : UDINT := 16#03B800;
  DFCid : UINT := 315;
  debounceMethod : USINT := TIME_UP_DOWN;
END_STRUCT;
END_TYPE

TYPE DFC_rbr_inK35OR : STRUCT
  DTC : UDINT := 16#03B700;
  DFCid : UINT := 314;
  debounceMethod : USINT := TIME_UP_DOWN;
END_STRUCT;
END_TYPE

TYPE DFC_rbr_inK34SCG : STRUCT
  DTC : UDINT := 16#03B600;
  DFCid : UINT := 313;
  debounceMethod : USINT := TIME_UP_DOWN;
END_STRUCT;
END_TYPE

TYPE DFC_rbr_inK34SCB : STRUCT
  DTC : UDINT := 16#03B500;
  DFCid : UINT := 312;
  debounceMethod : USINT := TIME_UP_DOWN;
END_STRUCT;
END_TYPE

TYPE DFC_rbr_inK34OR : STRUCT
  DTC : UDINT := 16#03B400;
  DFCid : UINT := 311;
  debounceMethod : USINT := TIME_UP_DOWN;
END_STRUCT;
END_TYPE

TYPE DFC_rbr_inK33SCG : STRUCT
  DTC : UDINT := 16#03B300;
  DFCid : UINT := 310;
  debounceMethod : USINT := TIME_UP_DOWN;
END_STRUCT;
END_TYPE

TYPE DFC_rbr_inK33SCB : STRUCT
  DTC : UDINT := 16#03B200;
  DFCid : UINT := 309;
  debounceMethod : USINT := TIME_UP_DOWN;
END_STRUCT;
END_TYPE

TYPE DFC_rbr_inK33OR : STRUCT
  DTC : UDINT := 16#03B100;
  DFCid : UINT := 308;
  debounceMethod : USINT := TIME_UP_DOWN;
END_STRUCT;
END_TYPE

TYPE DFC_rbr_inK32SCG : STRUCT
  DTC : UDINT := 16#03B000;
  DFCid : UINT := 307;
  debounceMethod : USINT := TIME_UP_DOWN;
END_STRUCT;
END_TYPE

TYPE DFC_rbr_inK32SCB : STRUCT
  DTC : UDINT := 16#03AF00;
  DFCid : UINT := 306;
  debounceMethod : USINT := TIME_UP_DOWN;
END_STRUCT;
END_TYPE

TYPE DFC_rbr_inK32OR : STRUCT
  DTC : UDINT := 16#03AE00;
  DFCid : UINT := 305;
  debounceMethod : USINT := TIME_UP_DOWN;
END_STRUCT;
END_TYPE

TYPE DFC_rbr_inK31SCG : STRUCT
  DTC : UDINT := 16#03AD00;
  DFCid : UINT := 304;
  debounceMethod : USINT := TIME_UP_DOWN;
END_STRUCT;
END_TYPE

TYPE DFC_rbr_inK31SCB : STRUCT
  DTC : UDINT := 16#03AC00;
  DFCid : UINT := 303;
  debounceMethod : USINT := TIME_UP_DOWN;
END_STRUCT;
END_TYPE

TYPE DFC_rbr_inK31OR : STRUCT
  DTC : UDINT := 16#03AB00;
  DFCid : UINT := 302;
  debounceMethod : USINT := TIME_UP_DOWN;
END_STRUCT;
END_TYPE

TYPE DFC_rbr_inK30ShuntSCB : STRUCT
  DTC : UDINT := 16#03AA00;
  DFCid : UINT := 301;
  debounceMethod : USINT := TIME_UP_DOWN;
END_STRUCT;
END_TYPE

TYPE DFC_rbr_inK30SCG : STRUCT
  DTC : UDINT := 16#03A900;
  DFCid : UINT := 300;
  debounceMethod : USINT := TIME_UP_DOWN;
END_STRUCT;
END_TYPE

TYPE DFC_rbr_inK30SCB : STRUCT
  DTC : UDINT := 16#03A800;
  DFCid : UINT := 299;
  debounceMethod : USINT := TIME_UP_DOWN;
END_STRUCT;
END_TYPE

TYPE DFC_rbr_inK30OR : STRUCT
  DTC : UDINT := 16#03A700;
  DFCid : UINT := 298;
  debounceMethod : USINT := TIME_UP_DOWN;
END_STRUCT;
END_TYPE

TYPE DFC_rbr_inK30AicSCG : STRUCT
  DTC : UDINT := 16#03A600;
  DFCid : UINT := 297;
  debounceMethod : USINT := TIME_UP_DOWN;
END_STRUCT;
END_TYPE

TYPE DFC_rbr_inK30AicSCB : STRUCT
  DTC : UDINT := 16#03A500;
  DFCid : UINT := 296;
  debounceMethod : USINT := TIME_UP_DOWN;
END_STRUCT;
END_TYPE

TYPE DFC_rbr_inK11SCG : STRUCT
  DTC : UDINT := 16#03A400;
  DFCid : UINT := 295;
  debounceMethod : USINT := TIME_UP_DOWN;
END_STRUCT;
END_TYPE

TYPE DFC_rbr_inK11SCB : STRUCT
  DTC : UDINT := 16#03A300;
  DFCid : UINT := 294;
  debounceMethod : USINT := TIME_UP_DOWN;
END_STRUCT;
END_TYPE

TYPE DFC_rbr_inK11OR : STRUCT
  DTC : UDINT := 16#03A200;
  DFCid : UINT := 293;
  debounceMethod : USINT := TIME_UP_DOWN;
END_STRUCT;
END_TYPE

TYPE DFC_rbr_inA59SCG : STRUCT
  DTC : UDINT := 16#135100;
  DFCid : UINT := 289;
  debounceMethod : USINT := TIME_UP_DOWN;
END_STRUCT;
END_TYPE

TYPE DFC_rbr_inA59SCB : STRUCT
  DTC : UDINT := 16#135000;
  DFCid : UINT := 288;
  debounceMethod : USINT := TIME_UP_DOWN;
END_STRUCT;
END_TYPE

TYPE DFC_rbr_inA59OL : STRUCT
  DTC : UDINT := 16#134F00;
  DFCid : UINT := 287;
  debounceMethod : USINT := TIME_UP_DOWN;
END_STRUCT;
END_TYPE

TYPE DFC_rbr_inA57SCG : STRUCT
  DTC : UDINT := 16#134E00;
  DFCid : UINT := 286;
  debounceMethod : USINT := TIME_UP_DOWN;
END_STRUCT;
END_TYPE

TYPE DFC_rbr_inA57SCB : STRUCT
  DTC : UDINT := 16#134D00;
  DFCid : UINT := 285;
  debounceMethod : USINT := TIME_UP_DOWN;
END_STRUCT;
END_TYPE

TYPE DFC_rbr_inA57OR : STRUCT
  DTC : UDINT := 16#134C00;
  DFCid : UINT := 284;
  debounceMethod : USINT := TIME_UP_DOWN;
END_STRUCT;
END_TYPE

TYPE DFC_rbr_inA44SCG : STRUCT
  DTC : UDINT := 16#134B00;
  DFCid : UINT := 283;
  debounceMethod : USINT := TIME_UP_DOWN;
END_STRUCT;
END_TYPE

TYPE DFC_rbr_inA44SCB : STRUCT
  DTC : UDINT := 16#134A00;
  DFCid : UINT := 282;
  debounceMethod : USINT := TIME_UP_DOWN;
END_STRUCT;
END_TYPE

TYPE DFC_rbr_inA44OL : STRUCT
  DTC : UDINT := 16#134900;
  DFCid : UINT := 281;
  debounceMethod : USINT := TIME_UP_DOWN;
END_STRUCT;
END_TYPE

TYPE DFC_rbr_inA43ShuntSCB : STRUCT
  DTC : UDINT := 16#134800;
  DFCid : UINT := 280;
  debounceMethod : USINT := TIME_UP_DOWN;
END_STRUCT;
END_TYPE

TYPE DFC_rbr_inA43SCG : STRUCT
  DTC : UDINT := 16#134700;
  DFCid : UINT := 279;
  debounceMethod : USINT := TIME_UP_DOWN;
END_STRUCT;
END_TYPE

TYPE DFC_rbr_inA43SCB : STRUCT
  DTC : UDINT := 16#134600;
  DFCid : UINT := 278;
  debounceMethod : USINT := TIME_UP_DOWN;
END_STRUCT;
END_TYPE

TYPE DFC_rbr_inA43OR : STRUCT
  DTC : UDINT := 16#134500;
  DFCid : UINT := 277;
  debounceMethod : USINT := TIME_UP_DOWN;
END_STRUCT;
END_TYPE

TYPE DFC_rbr_inA43AicSCG : STRUCT
  DTC : UDINT := 16#134400;
  DFCid : UINT := 276;
  debounceMethod : USINT := TIME_UP_DOWN;
END_STRUCT;
END_TYPE

TYPE DFC_rbr_inA43AicSCB : STRUCT
  DTC : UDINT := 16#134300;
  DFCid : UINT := 275;
  debounceMethod : USINT := TIME_UP_DOWN;
END_STRUCT;
END_TYPE

TYPE DFC_rbr_inA42SCG : STRUCT
  DTC : UDINT := 16#134200;
  DFCid : UINT := 274;
  debounceMethod : USINT := TIME_UP_DOWN;
END_STRUCT;
END_TYPE

TYPE DFC_rbr_inA42SCB : STRUCT
  DTC : UDINT := 16#134100;
  DFCid : UINT := 273;
  debounceMethod : USINT := TIME_UP_DOWN;
END_STRUCT;
END_TYPE

TYPE DFC_rbr_inA42OR : STRUCT
  DTC : UDINT := 16#134000;
  DFCid : UINT := 272;
  debounceMethod : USINT := TIME_UP_DOWN;
END_STRUCT;
END_TYPE

TYPE DFC_rbr_inA41SCG : STRUCT
  DTC : UDINT := 16#133F00;
  DFCid : UINT := 271;
  debounceMethod : USINT := TIME_UP_DOWN;
END_STRUCT;
END_TYPE

TYPE DFC_rbr_inA41SCB : STRUCT
  DTC : UDINT := 16#133E00;
  DFCid : UINT := 270;
  debounceMethod : USINT := TIME_UP_DOWN;
END_STRUCT;
END_TYPE

TYPE DFC_rbr_inA41OR : STRUCT
  DTC : UDINT := 16#133D00;
  DFCid : UINT := 269;
  debounceMethod : USINT := TIME_UP_DOWN;
END_STRUCT;
END_TYPE

TYPE DFC_rbr_inA40SCG : STRUCT
  DTC : UDINT := 16#133C00;
  DFCid : UINT := 268;
  debounceMethod : USINT := TIME_UP_DOWN;
END_STRUCT;
END_TYPE

TYPE DFC_rbr_inA40SCB : STRUCT
  DTC : UDINT := 16#133B00;
  DFCid : UINT := 267;
  debounceMethod : USINT := TIME_UP_DOWN;
END_STRUCT;
END_TYPE

TYPE DFC_rbr_inA40OR : STRUCT
  DTC : UDINT := 16#133A00;
  DFCid : UINT := 266;
  debounceMethod : USINT := TIME_UP_DOWN;
END_STRUCT;
END_TYPE

TYPE DFC_rbr_inA39ShuntSCB : STRUCT
  DTC : UDINT := 16#133900;
  DFCid : UINT := 265;
  debounceMethod : USINT := TIME_UP_DOWN;
END_STRUCT;
END_TYPE

TYPE DFC_rbr_inA39SCG : STRUCT
  DTC : UDINT := 16#133800;
  DFCid : UINT := 264;
  debounceMethod : USINT := TIME_UP_DOWN;
END_STRUCT;
END_TYPE

TYPE DFC_rbr_inA39SCB : STRUCT
  DTC : UDINT := 16#133700;
  DFCid : UINT := 263;
  debounceMethod : USINT := TIME_UP_DOWN;
END_STRUCT;
END_TYPE

TYPE DFC_rbr_inA39OR : STRUCT
  DTC : UDINT := 16#133600;
  DFCid : UINT := 262;
  debounceMethod : USINT := TIME_UP_DOWN;
END_STRUCT;
END_TYPE

TYPE DFC_rbr_inA39AicSCG : STRUCT
  DTC : UDINT := 16#133500;
  DFCid : UINT := 261;
  debounceMethod : USINT := TIME_UP_DOWN;
END_STRUCT;
END_TYPE

TYPE DFC_rbr_inA39AicSCB : STRUCT
  DTC : UDINT := 16#133400;
  DFCid : UINT := 260;
  debounceMethod : USINT := TIME_UP_DOWN;
END_STRUCT;
END_TYPE

TYPE DFC_rbr_inA38ShuntSCB : STRUCT
  DTC : UDINT := 16#133300;
  DFCid : UINT := 259;
  debounceMethod : USINT := TIME_UP_DOWN;
END_STRUCT;
END_TYPE

TYPE DFC_rbr_inA38SCG : STRUCT
  DTC : UDINT := 16#133200;
  DFCid : UINT := 258;
  debounceMethod : USINT := TIME_UP_DOWN;
END_STRUCT;
END_TYPE

TYPE DFC_rbr_inA38SCB : STRUCT
  DTC : UDINT := 16#133100;
  DFCid : UINT := 257;
  debounceMethod : USINT := TIME_UP_DOWN;
END_STRUCT;
END_TYPE

TYPE DFC_rbr_inA38OR : STRUCT
  DTC : UDINT := 16#133000;
  DFCid : UINT := 256;
  debounceMethod : USINT := TIME_UP_DOWN;
END_STRUCT;
END_TYPE

TYPE DFC_rbr_inA38AicSCG : STRUCT
  DTC : UDINT := 16#132F00;
  DFCid : UINT := 255;
  debounceMethod : USINT := TIME_UP_DOWN;
END_STRUCT;
END_TYPE

TYPE DFC_rbr_inA38AicSCB : STRUCT
  DTC : UDINT := 16#132E00;
  DFCid : UINT := 254;
  debounceMethod : USINT := TIME_UP_DOWN;
END_STRUCT;
END_TYPE

TYPE DFC_rbr_inA37ShuntSCB : STRUCT
  DTC : UDINT := 16#132D00;
  DFCid : UINT := 253;
  debounceMethod : USINT := TIME_UP_DOWN;
END_STRUCT;
END_TYPE

TYPE DFC_rbr_inA37SCG : STRUCT
  DTC : UDINT := 16#132C00;
  DFCid : UINT := 252;
  debounceMethod : USINT := TIME_UP_DOWN;
END_STRUCT;
END_TYPE

TYPE DFC_rbr_inA37SCB : STRUCT
  DTC : UDINT := 16#132B00;
  DFCid : UINT := 251;
  debounceMethod : USINT := TIME_UP_DOWN;
END_STRUCT;
END_TYPE

TYPE DFC_rbr_inA37OR : STRUCT
  DTC : UDINT := 16#132A00;
  DFCid : UINT := 250;
  debounceMethod : USINT := TIME_UP_DOWN;
END_STRUCT;
END_TYPE

TYPE DFC_rbr_inA37AicSCG : STRUCT
  DTC : UDINT := 16#132900;
  DFCid : UINT := 249;
  debounceMethod : USINT := TIME_UP_DOWN;
END_STRUCT;
END_TYPE

TYPE DFC_rbr_inA37AicSCB : STRUCT
  DTC : UDINT := 16#132800;
  DFCid : UINT := 248;
  debounceMethod : USINT := TIME_UP_DOWN;
END_STRUCT;
END_TYPE

TYPE DFC_rbr_inA36ShuntSCB : STRUCT
  DTC : UDINT := 16#132700;
  DFCid : UINT := 247;
  debounceMethod : USINT := TIME_UP_DOWN;
END_STRUCT;
END_TYPE

TYPE DFC_rbr_inA36SCG : STRUCT
  DTC : UDINT := 16#132600;
  DFCid : UINT := 246;
  debounceMethod : USINT := TIME_UP_DOWN;
END_STRUCT;
END_TYPE

TYPE DFC_rbr_inA36SCB : STRUCT
  DTC : UDINT := 16#132500;
  DFCid : UINT := 245;
  debounceMethod : USINT := TIME_UP_DOWN;
END_STRUCT;
END_TYPE

TYPE DFC_rbr_inA36OR : STRUCT
  DTC : UDINT := 16#132400;
  DFCid : UINT := 244;
  debounceMethod : USINT := TIME_UP_DOWN;
END_STRUCT;
END_TYPE

TYPE DFC_rbr_inA36AicSCG : STRUCT
  DTC : UDINT := 16#132300;
  DFCid : UINT := 243;
  debounceMethod : USINT := TIME_UP_DOWN;
END_STRUCT;
END_TYPE

TYPE DFC_rbr_inA36AicSCB : STRUCT
  DTC : UDINT := 16#132200;
  DFCid : UINT := 242;
  debounceMethod : USINT := TIME_UP_DOWN;
END_STRUCT;
END_TYPE

TYPE DFC_rbr_inA29SCG : STRUCT
  DTC : UDINT := 16#132100;
  DFCid : UINT := 241;
  debounceMethod : USINT := TIME_UP_DOWN;
END_STRUCT;
END_TYPE

TYPE DFC_rbr_inA29SCB : STRUCT
  DTC : UDINT := 16#132000;
  DFCid : UINT := 240;
  debounceMethod : USINT := TIME_UP_DOWN;
END_STRUCT;
END_TYPE

TYPE DFC_rbr_inA29OR : STRUCT
  DTC : UDINT := 16#131F00;
  DFCid : UINT := 239;
  debounceMethod : USINT := TIME_UP_DOWN;
END_STRUCT;
END_TYPE

TYPE DFC_rbr_inA28SCG : STRUCT
  DTC : UDINT := 16#131E00;
  DFCid : UINT := 238;
  debounceMethod : USINT := TIME_UP_DOWN;
END_STRUCT;
END_TYPE

TYPE DFC_rbr_inA28SCB : STRUCT
  DTC : UDINT := 16#131D00;
  DFCid : UINT := 237;
  debounceMethod : USINT := TIME_UP_DOWN;
END_STRUCT;
END_TYPE

TYPE DFC_rbr_inA28OR : STRUCT
  DTC : UDINT := 16#131C00;
  DFCid : UINT := 236;
  debounceMethod : USINT := TIME_UP_DOWN;
END_STRUCT;
END_TYPE

TYPE DFC_rbr_inA27SCG : STRUCT
  DTC : UDINT := 16#131B00;
  DFCid : UINT := 235;
  debounceMethod : USINT := TIME_UP_DOWN;
END_STRUCT;
END_TYPE

TYPE DFC_rbr_inA27SCB : STRUCT
  DTC : UDINT := 16#131A00;
  DFCid : UINT := 234;
  debounceMethod : USINT := TIME_UP_DOWN;
END_STRUCT;
END_TYPE

TYPE DFC_rbr_inA27OR : STRUCT
  DTC : UDINT := 16#131900;
  DFCid : UINT := 233;
  debounceMethod : USINT := TIME_UP_DOWN;
END_STRUCT;
END_TYPE

TYPE DFC_rbr_inA26SCG : STRUCT
  DTC : UDINT := 16#131800;
  DFCid : UINT := 232;
  debounceMethod : USINT := TIME_UP_DOWN;
END_STRUCT;
END_TYPE

TYPE DFC_rbr_inA26SCB : STRUCT
  DTC : UDINT := 16#131700;
  DFCid : UINT := 231;
  debounceMethod : USINT := TIME_UP_DOWN;
END_STRUCT;
END_TYPE

TYPE DFC_rbr_inA26OR : STRUCT
  DTC : UDINT := 16#131600;
  DFCid : UINT := 230;
  debounceMethod : USINT := TIME_UP_DOWN;
END_STRUCT;
END_TYPE

TYPE DFC_rbr_inA25SCG : STRUCT
  DTC : UDINT := 16#131500;
  DFCid : UINT := 229;
  debounceMethod : USINT := TIME_UP_DOWN;
END_STRUCT;
END_TYPE

TYPE DFC_rbr_inA25SCB : STRUCT
  DTC : UDINT := 16#131400;
  DFCid : UINT := 228;
  debounceMethod : USINT := TIME_UP_DOWN;
END_STRUCT;
END_TYPE

TYPE DFC_rbr_inA25OR : STRUCT
  DTC : UDINT := 16#131300;
  DFCid : UINT := 227;
  debounceMethod : USINT := TIME_UP_DOWN;
END_STRUCT;
END_TYPE

TYPE DFC_rbr_inA24SCG : STRUCT
  DTC : UDINT := 16#131200;
  DFCid : UINT := 226;
  debounceMethod : USINT := TIME_UP_DOWN;
END_STRUCT;
END_TYPE

TYPE DFC_rbr_inA24SCB : STRUCT
  DTC : UDINT := 16#131100;
  DFCid : UINT := 225;
  debounceMethod : USINT := TIME_UP_DOWN;
END_STRUCT;
END_TYPE

TYPE DFC_rbr_inA24OR : STRUCT
  DTC : UDINT := 16#131000;
  DFCid : UINT := 224;
  debounceMethod : USINT := TIME_UP_DOWN;
END_STRUCT;
END_TYPE

TYPE DFC_rbr_inA23SCG : STRUCT
  DTC : UDINT := 16#130F00;
  DFCid : UINT := 223;
  debounceMethod : USINT := TIME_UP_DOWN;
END_STRUCT;
END_TYPE

TYPE DFC_rbr_inA23SCB : STRUCT
  DTC : UDINT := 16#130E00;
  DFCid : UINT := 222;
  debounceMethod : USINT := TIME_UP_DOWN;
END_STRUCT;
END_TYPE

TYPE DFC_rbr_inA23OR : STRUCT
  DTC : UDINT := 16#130D00;
  DFCid : UINT := 221;
  debounceMethod : USINT := TIME_UP_DOWN;
END_STRUCT;
END_TYPE

TYPE DFC_rbr_inA22SCG : STRUCT
  DTC : UDINT := 16#130C00;
  DFCid : UINT := 220;
  debounceMethod : USINT := TIME_UP_DOWN;
END_STRUCT;
END_TYPE

TYPE DFC_rbr_inA22SCB : STRUCT
  DTC : UDINT := 16#130B00;
  DFCid : UINT := 219;
  debounceMethod : USINT := TIME_UP_DOWN;
END_STRUCT;
END_TYPE

TYPE DFC_rbr_inA22OR : STRUCT
  DTC : UDINT := 16#130A00;
  DFCid : UINT := 218;
  debounceMethod : USINT := TIME_UP_DOWN;
END_STRUCT;
END_TYPE

TYPE DFC_rbr_inA21SCG : STRUCT
  DTC : UDINT := 16#130900;
  DFCid : UINT := 217;
  debounceMethod : USINT := TIME_UP_DOWN;
END_STRUCT;
END_TYPE

TYPE DFC_rbr_inA21SCB : STRUCT
  DTC : UDINT := 16#130800;
  DFCid : UINT := 216;
  debounceMethod : USINT := TIME_UP_DOWN;
END_STRUCT;
END_TYPE

TYPE DFC_rbr_inA21OR : STRUCT
  DTC : UDINT := 16#130700;
  DFCid : UINT := 215;
  debounceMethod : USINT := TIME_UP_DOWN;
END_STRUCT;
END_TYPE

TYPE DFC_rbr_inA14SCG : STRUCT
  DTC : UDINT := 16#130600;
  DFCid : UINT := 214;
  debounceMethod : USINT := TIME_UP_DOWN;
END_STRUCT;
END_TYPE

TYPE DFC_rbr_inA14SCB : STRUCT
  DTC : UDINT := 16#130500;
  DFCid : UINT := 213;
  debounceMethod : USINT := TIME_UP_DOWN;
END_STRUCT;
END_TYPE

TYPE DFC_rbr_inA14OR : STRUCT
  DTC : UDINT := 16#130400;
  DFCid : UINT := 212;
  debounceMethod : USINT := TIME_UP_DOWN;
END_STRUCT;
END_TYPE

TYPE DFC_rbr_inA13SCG : STRUCT
  DTC : UDINT := 16#130300;
  DFCid : UINT := 211;
  debounceMethod : USINT := TIME_UP_DOWN;
END_STRUCT;
END_TYPE

TYPE DFC_rbr_inA13SCB : STRUCT
  DTC : UDINT := 16#130200;
  DFCid : UINT := 210;
  debounceMethod : USINT := TIME_UP_DOWN;
END_STRUCT;
END_TYPE

TYPE DFC_rbr_inA13OR : STRUCT
  DTC : UDINT := 16#130100;
  DFCid : UINT := 209;
  debounceMethod : USINT := TIME_UP_DOWN;
END_STRUCT;
END_TYPE

TYPE DFC_rbr_inK52SCB : STRUCT
  DTC : UDINT := 16#032600;
  DFCid : UINT := 372;
  debounceMethod : USINT := TIME_UP_DOWN;
END_STRUCT;
END_TYPE

TYPE DFC_rbr_inK52SCG : STRUCT
  DTC : UDINT := 16#032700;
  DFCid : UINT := 373;
  debounceMethod : USINT := TIME_UP_DOWN;
END_STRUCT;
END_TYPE

TYPE DFC_rbr_inK52OR : STRUCT
  DTC : UDINT := 16#032500;
  DFCid : UINT := 371;
  debounceMethod : USINT := TIME_UP_DOWN;
END_STRUCT;
END_TYPE

TYPE DFC_rbr_inK60SCB : STRUCT
  DTC : UDINT := 16#034400;
  DFCid : UINT := 402;
  debounceMethod : USINT := TIME_UP_DOWN;
END_STRUCT;
END_TYPE

TYPE DFC_rbr_inK60SCG : STRUCT
  DTC : UDINT := 16#034500;
  DFCid : UINT := 403;
  debounceMethod : USINT := TIME_UP_DOWN;
END_STRUCT;
END_TYPE

TYPE DFC_rbr_inK60OR : STRUCT
  DTC : UDINT := 16#034300;
  DFCid : UINT := 401;
  debounceMethod : USINT := TIME_UP_DOWN;
END_STRUCT;
END_TYPE

TYPE DFC_rbr_inK53SCB : STRUCT
  DTC : UDINT := 16#032900;
  DFCid : UINT := 375;
  debounceMethod : USINT := TIME_UP_DOWN;
END_STRUCT;
END_TYPE

TYPE DFC_rbr_inK53SCG : STRUCT
  DTC : UDINT := 16#032A00;
  DFCid : UINT := 376;
  debounceMethod : USINT := TIME_UP_DOWN;
END_STRUCT;
END_TYPE

TYPE DFC_rbr_inK53OR : STRUCT
  DTC : UDINT := 16#032800;
  DFCid : UINT := 374;
  debounceMethod : USINT := TIME_UP_DOWN;
END_STRUCT;
END_TYPE

TYPE DFC_rbr_inK59SCB : STRUCT
  DTC : UDINT := 16#034100;
  DFCid : UINT := 399;
  debounceMethod : USINT := TIME_UP_DOWN;
END_STRUCT;
END_TYPE

TYPE DFC_rbr_inK59SCG : STRUCT
  DTC : UDINT := 16#034200;
  DFCid : UINT := 400;
  debounceMethod : USINT := TIME_UP_DOWN;
END_STRUCT;
END_TYPE

TYPE DFC_rbr_inK59OR : STRUCT
  DTC : UDINT := 16#034000;
  DFCid : UINT := 398;
  debounceMethod : USINT := TIME_UP_DOWN;
END_STRUCT;
END_TYPE

TYPE DFC_rbr_inK39SCB : STRUCT
  DTC : UDINT := 16#031100;
  DFCid : UINT := 335;
  debounceMethod : USINT := TIME_UP_DOWN;
END_STRUCT;
END_TYPE

TYPE DFC_rbr_inK39SCG : STRUCT
  DTC : UDINT := 16#031200;
  DFCid : UINT := 336;
  debounceMethod : USINT := TIME_UP_DOWN;
END_STRUCT;
END_TYPE

TYPE DFC_rbr_inK39OR : STRUCT
  DTC : UDINT := 16#031000;
  DFCid : UINT := 334;
  debounceMethod : USINT := TIME_UP_DOWN;
END_STRUCT;
END_TYPE

TYPE DFC_rbr_inK38SCB : STRUCT
  DTC : UDINT := 16#030E00;
  DFCid : UINT := 329;
  debounceMethod : USINT := TIME_UP_DOWN;
END_STRUCT;
END_TYPE

TYPE DFC_rbr_inK38SCG : STRUCT
  DTC : UDINT := 16#030F00;
  DFCid : UINT := 330;
  debounceMethod : USINT := TIME_UP_DOWN;
END_STRUCT;
END_TYPE

TYPE DFC_rbr_inK38OR : STRUCT
  DTC : UDINT := 16#030D00;
  DFCid : UINT := 328;
  debounceMethod : USINT := TIME_UP_DOWN;
END_STRUCT;
END_TYPE

TYPE DFC_rbr_inK40SCB : STRUCT
  DTC : UDINT := 16#031400;
  DFCid : UINT := 341;
  debounceMethod : USINT := TIME_UP_DOWN;
END_STRUCT;
END_TYPE

TYPE DFC_rbr_inK40SCG : STRUCT
  DTC : UDINT := 16#031500;
  DFCid : UINT := 342;
  debounceMethod : USINT := TIME_UP_DOWN;
END_STRUCT;
END_TYPE

TYPE DFC_rbr_inK40OR : STRUCT
  DTC : UDINT := 16#031300;
  DFCid : UINT := 340;
  debounceMethod : USINT := TIME_UP_DOWN;
END_STRUCT;
END_TYPE

TYPE DFC_rbr_inK41SCB : STRUCT
  DTC : UDINT := 16#031700;
  DFCid : UINT := 347;
  debounceMethod : USINT := TIME_UP_DOWN;
END_STRUCT;
END_TYPE

TYPE DFC_rbr_inK41SCG : STRUCT
  DTC : UDINT := 16#031800;
  DFCid : UINT := 348;
  debounceMethod : USINT := TIME_UP_DOWN;
END_STRUCT;
END_TYPE

TYPE DFC_rbr_inK41OR : STRUCT
  DTC : UDINT := 16#031600;
  DFCid : UINT := 346;
  debounceMethod : USINT := TIME_UP_DOWN;
END_STRUCT;
END_TYPE

TYPE DFC_rbr_inK42SCB : STRUCT
  DTC : UDINT := 16#031A00;
  DFCid : UINT := 353;
  debounceMethod : USINT := TIME_UP_DOWN;
END_STRUCT;
END_TYPE

TYPE DFC_rbr_inK42SCG : STRUCT
  DTC : UDINT := 16#031B00;
  DFCid : UINT := 354;
  debounceMethod : USINT := TIME_UP_DOWN;
END_STRUCT;
END_TYPE

TYPE DFC_rbr_inK42OR : STRUCT
  DTC : UDINT := 16#031900;
  DFCid : UINT := 352;
  debounceMethod : USINT := TIME_UP_DOWN;
END_STRUCT;
END_TYPE

TYPE DFC_rbr_inK43SCB : STRUCT
  DTC : UDINT := 16#031D00;
  DFCid : UINT := 357;
  debounceMethod : USINT := TIME_UP_DOWN;
END_STRUCT;
END_TYPE

TYPE DFC_rbr_inK43SCG : STRUCT
  DTC : UDINT := 16#031E00;
  DFCid : UINT := 358;
  debounceMethod : USINT := TIME_UP_DOWN;
END_STRUCT;
END_TYPE

TYPE DFC_rbr_inK43OR : STRUCT
  DTC : UDINT := 16#031C00;
  DFCid : UINT := 356;
  debounceMethod : USINT := TIME_UP_DOWN;
END_STRUCT;
END_TYPE

TYPE DFC_rbr_inK54SCB : STRUCT
  DTC : UDINT := 16#032E00;
  DFCid : UINT := 380;
  debounceMethod : USINT := TIME_UP_DOWN;
END_STRUCT;
END_TYPE

TYPE DFC_rbr_inK54SCG : STRUCT
  DTC : UDINT := 16#032F00;
  DFCid : UINT := 381;
  debounceMethod : USINT := TIME_UP_DOWN;
END_STRUCT;
END_TYPE

TYPE DFC_rbr_inK54OR : STRUCT
  DTC : UDINT := 16#032D00;
  DFCid : UINT := 379;
  debounceMethod : USINT := TIME_UP_DOWN;
END_STRUCT;
END_TYPE

TYPE DFC_rbr_inK55SCB : STRUCT
  DTC : UDINT := 16#033400;
  DFCid : UINT := 386;
  debounceMethod : USINT := TIME_UP_DOWN;
END_STRUCT;
END_TYPE

TYPE DFC_rbr_inK55SCG : STRUCT
  DTC : UDINT := 16#033500;
  DFCid : UINT := 387;
  debounceMethod : USINT := TIME_UP_DOWN;
END_STRUCT;
END_TYPE

TYPE DFC_rbr_inK55OR : STRUCT
  DTC : UDINT := 16#033300;
  DFCid : UINT := 385;
  debounceMethod : USINT := TIME_UP_DOWN;
END_STRUCT;
END_TYPE

TYPE DFC_rbr_inK57SCB : STRUCT
  DTC : UDINT := 16#033B00;
  DFCid : UINT := 393;
  debounceMethod : USINT := TIME_UP_DOWN;
END_STRUCT;
END_TYPE

TYPE DFC_rbr_inK57SCG : STRUCT
  DTC : UDINT := 16#033C00;
  DFCid : UINT := 394;
  debounceMethod : USINT := TIME_UP_DOWN;
END_STRUCT;
END_TYPE

TYPE DFC_rbr_inK57OR : STRUCT
  DTC : UDINT := 16#033A00;
  DFCid : UINT := 392;
  debounceMethod : USINT := TIME_UP_DOWN;
END_STRUCT;
END_TYPE

TYPE DFC_rbr_inK58SCB : STRUCT
  DTC : UDINT := 16#033E00;
  DFCid : UINT := 396;
  debounceMethod : USINT := TIME_UP_DOWN;
END_STRUCT;
END_TYPE

TYPE DFC_rbr_inK58SCG : STRUCT
  DTC : UDINT := 16#033F00;
  DFCid : UINT := 397;
  debounceMethod : USINT := TIME_UP_DOWN;
END_STRUCT;
END_TYPE

TYPE DFC_rbr_inK58OR : STRUCT
  DTC : UDINT := 16#033D00;
  DFCid : UINT := 395;
  debounceMethod : USINT := TIME_UP_DOWN;
END_STRUCT;
END_TYPE

TYPE DFC_rbr_inK36SCB : STRUCT
  DTC : UDINT := 16#030500;
  DFCid : UINT := 318;
  debounceMethod : USINT := TIME_UP_DOWN;
END_STRUCT;
END_TYPE

TYPE DFC_rbr_inK36SCG : STRUCT
  DTC : UDINT := 16#030600;
  DFCid : UINT := 319;
  debounceMethod : USINT := TIME_UP_DOWN;
END_STRUCT;
END_TYPE

TYPE DFC_rbr_inK36OR : STRUCT
  DTC : UDINT := 16#030400;
  DFCid : UINT := 317;
  debounceMethod : USINT := TIME_UP_DOWN;
END_STRUCT;
END_TYPE

TYPE DFC_rbr_inK56SCB : STRUCT
  DTC : UDINT := 16#033800;
  DFCid : UINT := 390;
  debounceMethod : USINT := TIME_UP_DOWN;
END_STRUCT;
END_TYPE

TYPE DFC_rbr_inK56SCG : STRUCT
  DTC : UDINT := 16#033900;
  DFCid : UINT := 391;
  debounceMethod : USINT := TIME_UP_DOWN;
END_STRUCT;
END_TYPE

TYPE DFC_rbr_inK56OR : STRUCT
  DTC : UDINT := 16#033700;
  DFCid : UINT := 389;
  debounceMethod : USINT := TIME_UP_DOWN;
END_STRUCT;
END_TYPE

TYPE DFC_rbr_inK45SCB : STRUCT
  DTC : UDINT := 16#032300;
  DFCid : UINT := 368;
  debounceMethod : USINT := TIME_UP_DOWN;
END_STRUCT;
END_TYPE

TYPE DFC_rbr_inK45SCG : STRUCT
  DTC : UDINT := 16#032400;
  DFCid : UINT := 369;
  debounceMethod : USINT := TIME_UP_DOWN;
END_STRUCT;
END_TYPE

TYPE DFC_rbr_inK45OR : STRUCT
  DTC : UDINT := 16#032200;
  DFCid : UINT := 367;
  debounceMethod : USINT := TIME_UP_DOWN;
END_STRUCT;
END_TYPE

TYPE DFC_rbr_inK44SCB : STRUCT
  DTC : UDINT := 16#032000;
  DFCid : UINT := 362;
  debounceMethod : USINT := TIME_UP_DOWN;
END_STRUCT;
END_TYPE

TYPE DFC_rbr_inK44SCG : STRUCT
  DTC : UDINT := 16#032100;
  DFCid : UINT := 363;
  debounceMethod : USINT := TIME_UP_DOWN;
END_STRUCT;
END_TYPE

TYPE DFC_rbr_inK44OR : STRUCT
  DTC : UDINT := 16#031F00;
  DFCid : UINT := 361;
  debounceMethod : USINT := TIME_UP_DOWN;
END_STRUCT;
END_TYPE

TYPE DFC_rbr_inK65SCB : STRUCT
  DTC : UDINT := 16#035600;
  DFCid : UINT := 428;
  debounceMethod : USINT := TIME_UP_DOWN;
END_STRUCT;
END_TYPE

TYPE DFC_rbr_inK65SCG : STRUCT
  DTC : UDINT := 16#035700;
  DFCid : UINT := 429;
  debounceMethod : USINT := TIME_UP_DOWN;
END_STRUCT;
END_TYPE

TYPE DFC_rbr_inK65OR : STRUCT
  DTC : UDINT := 16#035500;
  DFCid : UINT := 427;
  debounceMethod : USINT := TIME_UP_DOWN;
END_STRUCT;
END_TYPE

TYPE DFC_rbr_inK63SCB : STRUCT
  DTC : UDINT := 16#035000;
  DFCid : UINT := 416;
  debounceMethod : USINT := TIME_UP_DOWN;
END_STRUCT;
END_TYPE

TYPE DFC_rbr_inK63SCG : STRUCT
  DTC : UDINT := 16#035100;
  DFCid : UINT := 417;
  debounceMethod : USINT := TIME_UP_DOWN;
END_STRUCT;
END_TYPE

TYPE DFC_rbr_inK63OR : STRUCT
  DTC : UDINT := 16#034F00;
  DFCid : UINT := 415;
  debounceMethod : USINT := TIME_UP_DOWN;
END_STRUCT;
END_TYPE

TYPE DFC_rbr_inK64SCB : STRUCT
  DTC : UDINT := 16#035300;
  DFCid : UINT := 422;
  debounceMethod : USINT := TIME_UP_DOWN;
END_STRUCT;
END_TYPE

TYPE DFC_rbr_inK64SCG : STRUCT
  DTC : UDINT := 16#035400;
  DFCid : UINT := 423;
  debounceMethod : USINT := TIME_UP_DOWN;
END_STRUCT;
END_TYPE

TYPE DFC_rbr_inK64OR : STRUCT
  DTC : UDINT := 16#035200;
  DFCid : UINT := 421;
  debounceMethod : USINT := TIME_UP_DOWN;
END_STRUCT;
END_TYPE

TYPE DFC_rbr_inK62SCB : STRUCT
  DTC : UDINT := 16#034D00;
  DFCid : UINT := 411;
  debounceMethod : USINT := TIME_UP_DOWN;
END_STRUCT;
END_TYPE

TYPE DFC_rbr_inK62SCG : STRUCT
  DTC : UDINT := 16#034E00;
  DFCid : UINT := 412;
  debounceMethod : USINT := TIME_UP_DOWN;
END_STRUCT;
END_TYPE

TYPE DFC_rbr_inK62OR : STRUCT
  DTC : UDINT := 16#034C00;
  DFCid : UINT := 410;
  debounceMethod : USINT := TIME_UP_DOWN;
END_STRUCT;
END_TYPE

TYPE DFC_rbr_inK37SCB : STRUCT
  DTC : UDINT := 16#030A00;
  DFCid : UINT := 323;
  debounceMethod : USINT := TIME_UP_DOWN;
END_STRUCT;
END_TYPE

TYPE DFC_rbr_inK37SCG : STRUCT
  DTC : UDINT := 16#030B00;
  DFCid : UINT := 324;
  debounceMethod : USINT := TIME_UP_DOWN;
END_STRUCT;
END_TYPE

TYPE DFC_rbr_inK37OR : STRUCT
  DTC : UDINT := 16#030900;
  DFCid : UINT := 322;
  debounceMethod : USINT := TIME_UP_DOWN;
END_STRUCT;
END_TYPE

TYPE DFC_rbr_inK61SCB : STRUCT
  DTC : UDINT := 16#034900;
  DFCid : UINT := 407;
  debounceMethod : USINT := TIME_UP_DOWN;
END_STRUCT;
END_TYPE

TYPE DFC_rbr_inK61SCG : STRUCT
  DTC : UDINT := 16#034A00;
  DFCid : UINT := 408;
  debounceMethod : USINT := TIME_UP_DOWN;
END_STRUCT;
END_TYPE

TYPE DFC_rbr_inK61OR : STRUCT
  DTC : UDINT := 16#034800;
  DFCid : UINT := 406;
  debounceMethod : USINT := TIME_UP_DOWN;
END_STRUCT;
END_TYPE

TYPE DFC_rbr_inK78SCB : STRUCT
  DTC : UDINT := 16#036500;
  DFCid : UINT := 444;
  debounceMethod : USINT := TIME_UP_DOWN;
END_STRUCT;
END_TYPE

TYPE DFC_rbr_inK78SCG : STRUCT
  DTC : UDINT := 16#036600;
  DFCid : UINT := 445;
  debounceMethod : USINT := TIME_UP_DOWN;
END_STRUCT;
END_TYPE

TYPE DFC_rbr_inK78OR : STRUCT
  DTC : UDINT := 16#036400;
  DFCid : UINT := 443;
  debounceMethod : USINT := TIME_UP_DOWN;
END_STRUCT;
END_TYPE

TYPE DFC_rbr_inK76SCB : STRUCT
  DTC : UDINT := 16#035F00;
  DFCid : UINT := 438;
  debounceMethod : USINT := TIME_UP_DOWN;
END_STRUCT;
END_TYPE

TYPE DFC_rbr_inK76SCG : STRUCT
  DTC : UDINT := 16#036000;
  DFCid : UINT := 439;
  debounceMethod : USINT := TIME_UP_DOWN;
END_STRUCT;
END_TYPE

TYPE DFC_rbr_inK76OR : STRUCT
  DTC : UDINT := 16#035E00;
  DFCid : UINT := 437;
  debounceMethod : USINT := TIME_UP_DOWN;
END_STRUCT;
END_TYPE

TYPE DFC_rbr_inK74SCB : STRUCT
  DTC : UDINT := 16#035900;
  DFCid : UINT := 432;
  debounceMethod : USINT := TIME_UP_DOWN;
END_STRUCT;
END_TYPE

TYPE DFC_rbr_inK74SCG : STRUCT
  DTC : UDINT := 16#035A00;
  DFCid : UINT := 433;
  debounceMethod : USINT := TIME_UP_DOWN;
END_STRUCT;
END_TYPE

TYPE DFC_rbr_inK74OR : STRUCT
  DTC : UDINT := 16#035800;
  DFCid : UINT := 431;
  debounceMethod : USINT := TIME_UP_DOWN;
END_STRUCT;
END_TYPE

TYPE DFC_rbr_inK77SCB : STRUCT
  DTC : UDINT := 16#036200;
  DFCid : UINT := 441;
  debounceMethod : USINT := TIME_UP_DOWN;
END_STRUCT;
END_TYPE

TYPE DFC_rbr_inK77SCG : STRUCT
  DTC : UDINT := 16#036300;
  DFCid : UINT := 442;
  debounceMethod : USINT := TIME_UP_DOWN;
END_STRUCT;
END_TYPE

TYPE DFC_rbr_inK77OR : STRUCT
  DTC : UDINT := 16#036100;
  DFCid : UINT := 440;
  debounceMethod : USINT := TIME_UP_DOWN;
END_STRUCT;
END_TYPE

TYPE DFC_rbr_inK10SCB : STRUCT
  DTC : UDINT := 16#030200;
  DFCid : UINT := 291;
  debounceMethod : USINT := TIME_UP_DOWN;
END_STRUCT;
END_TYPE

TYPE DFC_rbr_inK10SCG : STRUCT
  DTC : UDINT := 16#030300;
  DFCid : UINT := 292;
  debounceMethod : USINT := TIME_UP_DOWN;
END_STRUCT;
END_TYPE

TYPE DFC_rbr_inK10OR : STRUCT
  DTC : UDINT := 16#030100;
  DFCid : UINT := 290;
  debounceMethod : USINT := TIME_UP_DOWN;
END_STRUCT;
END_TYPE

TYPE DFC_rbr_inK75SCB : STRUCT
  DTC : UDINT := 16#035C00;
  DFCid : UINT := 435;
  debounceMethod : USINT := TIME_UP_DOWN;
END_STRUCT;
END_TYPE

TYPE DFC_rbr_inK75SCG : STRUCT
  DTC : UDINT := 16#035D00;
  DFCid : UINT := 436;
  debounceMethod : USINT := TIME_UP_DOWN;
END_STRUCT;
END_TYPE

TYPE DFC_rbr_inK75OR : STRUCT
  DTC : UDINT := 16#035B00;
  DFCid : UINT := 434;
  debounceMethod : USINT := TIME_UP_DOWN;
END_STRUCT;
END_TYPE

TYPE DFC_rbr_inK54AicSCB : STRUCT
  DTC : UDINT := 16#032B00;
  DFCid : UINT := 377;
  debounceMethod : USINT := TIME_UP_DOWN;
END_STRUCT;
END_TYPE

TYPE DFC_rbr_inK54AicSCG : STRUCT
  DTC : UDINT := 16#032C00;
  DFCid : UINT := 378;
  debounceMethod : USINT := TIME_UP_DOWN;
END_STRUCT;
END_TYPE

TYPE DFC_rbr_inK55AicSCB : STRUCT
  DTC : UDINT := 16#033100;
  DFCid : UINT := 383;
  debounceMethod : USINT := TIME_UP_DOWN;
END_STRUCT;
END_TYPE

TYPE DFC_rbr_inK55AicSCG : STRUCT
  DTC : UDINT := 16#033200;
  DFCid : UINT := 384;
  debounceMethod : USINT := TIME_UP_DOWN;
END_STRUCT;
END_TYPE

TYPE DFC_rbr_inK37AicSCB : STRUCT
  DTC : UDINT := 16#030700;
  DFCid : UINT := 320;
  debounceMethod : USINT := TIME_UP_DOWN;
END_STRUCT;
END_TYPE

TYPE DFC_rbr_inK37AicSCG : STRUCT
  DTC : UDINT := 16#030800;
  DFCid : UINT := 321;
  debounceMethod : USINT := TIME_UP_DOWN;
END_STRUCT;
END_TYPE

TYPE DFC_rbr_inK61AicSCB : STRUCT
  DTC : UDINT := 16#034600;
  DFCid : UINT := 404;
  debounceMethod : USINT := TIME_UP_DOWN;
END_STRUCT;
END_TYPE

TYPE DFC_rbr_inK61AicSCG : STRUCT
  DTC : UDINT := 16#034700;
  DFCid : UINT := 405;
  debounceMethod : USINT := TIME_UP_DOWN;
END_STRUCT;
END_TYPE

TYPE DFC_rbr_inK54ShuntSCB : STRUCT
  DTC : UDINT := 16#033000;
  DFCid : UINT := 382;
  debounceMethod : USINT := TIME_UP_DOWN;
END_STRUCT;
END_TYPE

TYPE DFC_rbr_inK55ShuntSCB : STRUCT
  DTC : UDINT := 16#033600;
  DFCid : UINT := 388;
  debounceMethod : USINT := TIME_UP_DOWN;
END_STRUCT;
END_TYPE

TYPE DFC_rbr_inK37ShuntSCB : STRUCT
  DTC : UDINT := 16#030C00;
  DFCid : UINT := 325;
  debounceMethod : USINT := TIME_UP_DOWN;
END_STRUCT;
END_TYPE

TYPE DFC_rbr_inK61ShuntSCB : STRUCT
  DTC : UDINT := 16#034B00;
  DFCid : UINT := 409;
  debounceMethod : USINT := TIME_UP_DOWN;
END_STRUCT;
END_TYPE

TYPE DFC_rbr_inDi : STRUCT
  DTC : UDINT := 16#038700;
  DFCid : UINT := 891;
  debounceMethod : USINT := NO_DEBOUNCE;
END_STRUCT;
END_TYPE

TYPE DFC_rbr_inAi : STRUCT
  DTC : UDINT := 16#038000;
  DFCid : UINT := 882;
  debounceMethod : USINT := NO_DEBOUNCE;
END_STRUCT;
END_TYPE

TYPE DFC_rbr_inAiv : STRUCT
  DTC : UDINT := 16#038500;
  DFCid : UINT := 888;
  debounceMethod : USINT := NO_DEBOUNCE;
END_STRUCT;
END_TYPE

TYPE DFC_rbr_inAid : STRUCT
  DTC : UDINT := 16#038300;
  DFCid : UINT := 886;
  debounceMethod : USINT := NO_DEBOUNCE;
END_STRUCT;
END_TYPE

TYPE DFC_rbr_inAic : STRUCT
  DTC : UDINT := 16#038100;
  DFCid : UINT := 883;
  debounceMethod : USINT := NO_DEBOUNCE;
END_STRUCT;
END_TYPE

TYPE DFC_rbr_inRi : STRUCT
  DTC : UDINT := 16#038A00;
  DFCid : UINT := 899;
  debounceMethod : USINT := NO_DEBOUNCE;
END_STRUCT;
END_TYPE

TYPE DFC_rbr_inFiCfg : STRUCT
  DTC : UDINT := 16#038900;
  DFCid : UINT := 893;
  debounceMethod : USINT := NO_DEBOUNCE;
END_STRUCT;
END_TYPE

TYPE DFC_rbr_inFi : STRUCT
  DTC : UDINT := 16#038800;
  DFCid : UINT := 892;
  debounceMethod : USINT := NO_DEBOUNCE;
END_STRUCT;
END_TYPE

TYPE DFC_rbr_inAivCfg : STRUCT
  DTC : UDINT := 16#038600;
  DFCid : UINT := 889;
  debounceMethod : USINT := NO_DEBOUNCE;
END_STRUCT;
END_TYPE

TYPE DFC_rbr_inAidCfg : STRUCT
  DTC : UDINT := 16#038400;
  DFCid : UINT := 887;
  debounceMethod : USINT := NO_DEBOUNCE;
END_STRUCT;
END_TYPE

TYPE DFC_rbr_inAicCfg : STRUCT
  DTC : UDINT := 16#038200;
  DFCid : UINT := 884;
  debounceMethod : USINT := NO_DEBOUNCE;
END_STRUCT;
END_TYPE

TYPE DFC_rbr_inAicGetStatus : STRUCT
  DTC : UDINT := 16#038D00;
  DFCid : UINT := 885;
  debounceMethod : USINT := NO_DEBOUNCE;
END_STRUCT;
END_TYPE

TYPE DFC_rbr_inRiGetStatus : STRUCT
  DTC : UDINT := 16#038E00;
  DFCid : UINT := 902;
  debounceMethod : USINT := NO_DEBOUNCE;
END_STRUCT;
END_TYPE

TYPE DFC_rbr_inFiGetStatus : STRUCT
  DTC : UDINT := 16#038F00;
  DFCid : UINT := 894;
  debounceMethod : USINT := NO_DEBOUNCE;
END_STRUCT;
END_TYPE

TYPE DFC_rbr_inSentEnable : STRUCT
  DTC : UDINT := 16#039000;
  DFCid : UINT := 906;
  debounceMethod : USINT := NO_DEBOUNCE;
END_STRUCT;
END_TYPE

TYPE DFC_rbr_inSentDisable : STRUCT
  DTC : UDINT := 16#039100;
  DFCid : UINT := 905;
  debounceMethod : USINT := NO_DEBOUNCE;
END_STRUCT;
END_TYPE

TYPE DFC_rbr_inSentGetFD : STRUCT
  DTC : UDINT := 16#039200;
  DFCid : UINT := 908;
  debounceMethod : USINT := NO_DEBOUNCE;
END_STRUCT;
END_TYPE

TYPE DFC_rbr_inSentGetSD : STRUCT
  DTC : UDINT := 16#039300;
  DFCid : UINT := 909;
  debounceMethod : USINT := NO_DEBOUNCE;
END_STRUCT;
END_TYPE

TYPE DFC_rbr_inSentGetStatus : STRUCT
  DTC : UDINT := 16#039400;
  DFCid : UINT := 911;
  debounceMethod : USINT := NO_DEBOUNCE;
END_STRUCT;
END_TYPE

TYPE DFC_rbr_inSentGetErrorStatus : STRUCT
  DTC : UDINT := 16#039500;
  DFCid : UINT := 907;
  debounceMethod : USINT := NO_DEBOUNCE;
END_STRUCT;
END_TYPE

TYPE DFC_rbr_inSentRegisterFDFifo : STRUCT
  DTC : UDINT := 16#039600;
  DFCid : UINT := 914;
  debounceMethod : USINT := NO_DEBOUNCE;
END_STRUCT;
END_TYPE

TYPE DFC_rbr_inSentRegisterCopyFDFifo : STRUCT
  DTC : UDINT := 16#039700;
  DFCid : UINT := 913;
  debounceMethod : USINT := NO_DEBOUNCE;
END_STRUCT;
END_TYPE

TYPE DFC_rbr_inSentCopyFDFifo : STRUCT
  DTC : UDINT := 16#039800;
  DFCid : UINT := 904;
  debounceMethod : USINT := NO_DEBOUNCE;
END_STRUCT;
END_TYPE

TYPE DFC_rbr_inSentRegisterSDDataboxes : STRUCT
  DTC : UDINT := 16#039900;
  DFCid : UINT := 915;
  debounceMethod : USINT := NO_DEBOUNCE;
END_STRUCT;
END_TYPE

TYPE DFC_rbr_inSentInitSDDatabox : STRUCT
  DTC : UDINT := 16#039A00;
  DFCid : UINT := 912;
  debounceMethod : USINT := NO_DEBOUNCE;
END_STRUCT;
END_TYPE

TYPE DFC_rbr_inSentGetSDDatabox : STRUCT
  DTC : UDINT := 16#039B00;
  DFCid : UINT := 910;
  debounceMethod : USINT := NO_DEBOUNCE;
END_STRUCT;
END_TYPE

TYPE DFC_rbr_inAivGetStatus : STRUCT
  DTC : UDINT := 16#038C00;
  DFCid : UINT := 890;
  debounceMethod : USINT := NO_DEBOUNCE;
END_STRUCT;
END_TYPE

TYPE DFC_rbr_inRiCfg : STRUCT
  DTC : UDINT := 16#038B00;
  DFCid : UINT := 900;
  debounceMethod : USINT := NO_DEBOUNCE;
END_STRUCT;
END_TYPE

TYPE DFC_rbr_inRiCfgTemp : STRUCT
  DTC : UDINT := 16#039C00;
  DFCid : UINT := 901;
  debounceMethod : USINT := NO_DEBOUNCE;
END_STRUCT;
END_TYPE

TYPE DFC_rbr_inRiGetTemp : STRUCT
  DTC : UDINT := 16#039D00;
  DFCid : UINT := 903;
  debounceMethod : USINT := NO_DEBOUNCE;
END_STRUCT;
END_TYPE

TYPE DFC_rbr_outK16SCB : STRUCT
  DTC : UDINT := 16#042A00;
  DFCid : UINT := 661;
  debounceMethod : USINT := TIME_UP_DOWN;
END_STRUCT;
END_TYPE

TYPE DFC_rbr_outK16SCG : STRUCT
  DTC : UDINT := 16#042B00;
  DFCid : UINT := 662;
  debounceMethod : USINT := TIME_UP_DOWN;
END_STRUCT;
END_TYPE

TYPE DFC_rbr_outK16OL : STRUCT
  DTC : UDINT := 16#042800;
  DFCid : UINT := 658;
  debounceMethod : USINT := TIME_UP_DOWN;
END_STRUCT;
END_TYPE

TYPE DFC_rbr_outK16OC : STRUCT
  DTC : UDINT := 16#042700;
  DFCid : UINT := 1045;
  debounceMethod : USINT := NO_DEBOUNCE;
END_STRUCT;
END_TYPE

TYPE DFC_rbr_outK16OT : STRUCT
  DTC : UDINT := 16#042900;
  DFCid : UINT := 660;
  debounceMethod : USINT := TIME_UP_DOWN;
END_STRUCT;
END_TYPE

TYPE DFC_rbr_outK15SCB : STRUCT
  DTC : UDINT := 16#042500;
  DFCid : UINT := 656;
  debounceMethod : USINT := TIME_UP_DOWN;
END_STRUCT;
END_TYPE

TYPE DFC_rbr_outK15SCG : STRUCT
  DTC : UDINT := 16#042600;
  DFCid : UINT := 657;
  debounceMethod : USINT := TIME_UP_DOWN;
END_STRUCT;
END_TYPE

TYPE DFC_rbr_outK15OL : STRUCT
  DTC : UDINT := 16#042300;
  DFCid : UINT := 653;
  debounceMethod : USINT := TIME_UP_DOWN;
END_STRUCT;
END_TYPE

TYPE DFC_rbr_outK15OC : STRUCT
  DTC : UDINT := 16#042200;
  DFCid : UINT := 1043;
  debounceMethod : USINT := NO_DEBOUNCE;
END_STRUCT;
END_TYPE

TYPE DFC_rbr_outK15OT : STRUCT
  DTC : UDINT := 16#042400;
  DFCid : UINT := 655;
  debounceMethod : USINT := TIME_UP_DOWN;
END_STRUCT;
END_TYPE

TYPE DFC_rbr_outK13SCB : STRUCT
  DTC : UDINT := 16#041B00;
  DFCid : UINT := 646;
  debounceMethod : USINT := TIME_UP_DOWN;
END_STRUCT;
END_TYPE

TYPE DFC_rbr_outK13SCG : STRUCT
  DTC : UDINT := 16#041C00;
  DFCid : UINT := 647;
  debounceMethod : USINT := TIME_UP_DOWN;
END_STRUCT;
END_TYPE

TYPE DFC_rbr_outK13OL : STRUCT
  DTC : UDINT := 16#041900;
  DFCid : UINT := 644;
  debounceMethod : USINT := TIME_UP_DOWN;
END_STRUCT;
END_TYPE

TYPE DFC_rbr_outK13OC : STRUCT
  DTC : UDINT := 16#041800;
  DFCid : UINT := 1039;
  debounceMethod : USINT := NO_DEBOUNCE;
END_STRUCT;
END_TYPE

TYPE DFC_rbr_outK13OT : STRUCT
  DTC : UDINT := 16#041A00;
  DFCid : UINT := 645;
  debounceMethod : USINT := TIME_UP_DOWN;
END_STRUCT;
END_TYPE

TYPE DFC_rbr_outK12SCB : STRUCT
  DTC : UDINT := 16#041600;
  DFCid : UINT := 642;
  debounceMethod : USINT := TIME_UP_DOWN;
END_STRUCT;
END_TYPE

TYPE DFC_rbr_outK12SCG : STRUCT
  DTC : UDINT := 16#041700;
  DFCid : UINT := 643;
  debounceMethod : USINT := TIME_UP_DOWN;
END_STRUCT;
END_TYPE

TYPE DFC_rbr_outK12OL : STRUCT
  DTC : UDINT := 16#041400;
  DFCid : UINT := 640;
  debounceMethod : USINT := TIME_UP_DOWN;
END_STRUCT;
END_TYPE

TYPE DFC_rbr_outK12OC : STRUCT
  DTC : UDINT := 16#041300;
  DFCid : UINT := 1037;
  debounceMethod : USINT := NO_DEBOUNCE;
END_STRUCT;
END_TYPE

TYPE DFC_rbr_outK12OT : STRUCT
  DTC : UDINT := 16#041500;
  DFCid : UINT := 641;
  debounceMethod : USINT := TIME_UP_DOWN;
END_STRUCT;
END_TYPE

TYPE DFC_rbr_outK84SCB : STRUCT
  DTC : UDINT := 16#045500;
  DFCid : UINT := 706;
  debounceMethod : USINT := TIME_UP_DOWN;
END_STRUCT;
END_TYPE

TYPE DFC_rbr_outK84SCG : STRUCT
  DTC : UDINT := 16#045600;
  DFCid : UINT := 707;
  debounceMethod : USINT := TIME_UP_DOWN;
END_STRUCT;
END_TYPE

TYPE DFC_rbr_outK84OL : STRUCT
  DTC : UDINT := 16#045300;
  DFCid : UINT := 704;
  debounceMethod : USINT := TIME_UP_DOWN;
END_STRUCT;
END_TYPE

TYPE DFC_rbr_outK84OT : STRUCT
  DTC : UDINT := 16#045400;
  DFCid : UINT := 705;
  debounceMethod : USINT := TIME_UP_DOWN;
END_STRUCT;
END_TYPE

TYPE DFC_rbr_outK85SCB : STRUCT
  DTC : UDINT := 16#045900;
  DFCid : UINT := 710;
  debounceMethod : USINT := TIME_UP_DOWN;
END_STRUCT;
END_TYPE

TYPE DFC_rbr_outK85SCG : STRUCT
  DTC : UDINT := 16#045A00;
  DFCid : UINT := 711;
  debounceMethod : USINT := TIME_UP_DOWN;
END_STRUCT;
END_TYPE

TYPE DFC_rbr_outK85OT : STRUCT
  DTC : UDINT := 16#045800;
  DFCid : UINT := 709;
  debounceMethod : USINT := TIME_UP_DOWN;
END_STRUCT;
END_TYPE

TYPE DFC_rbr_outK85OL : STRUCT
  DTC : UDINT := 16#045700;
  DFCid : UINT := 708;
  debounceMethod : USINT := TIME_UP_DOWN;
END_STRUCT;
END_TYPE

TYPE DFC_rbr_outK86SCB : STRUCT
  DTC : UDINT := 16#045D00;
  DFCid : UINT := 714;
  debounceMethod : USINT := TIME_UP_DOWN;
END_STRUCT;
END_TYPE

TYPE DFC_rbr_outK86SCG : STRUCT
  DTC : UDINT := 16#045E00;
  DFCid : UINT := 715;
  debounceMethod : USINT := TIME_UP_DOWN;
END_STRUCT;
END_TYPE

TYPE DFC_rbr_outK86OL : STRUCT
  DTC : UDINT := 16#045B00;
  DFCid : UINT := 712;
  debounceMethod : USINT := TIME_UP_DOWN;
END_STRUCT;
END_TYPE

TYPE DFC_rbr_outK86OT : STRUCT
  DTC : UDINT := 16#045C00;
  DFCid : UINT := 713;
  debounceMethod : USINT := TIME_UP_DOWN;
END_STRUCT;
END_TYPE

TYPE DFC_rbr_outK87SCB : STRUCT
  DTC : UDINT := 16#046100;
  DFCid : UINT := 718;
  debounceMethod : USINT := TIME_UP_DOWN;
END_STRUCT;
END_TYPE

TYPE DFC_rbr_outK87SCG : STRUCT
  DTC : UDINT := 16#046200;
  DFCid : UINT := 719;
  debounceMethod : USINT := TIME_UP_DOWN;
END_STRUCT;
END_TYPE

TYPE DFC_rbr_outK87OL : STRUCT
  DTC : UDINT := 16#045F00;
  DFCid : UINT := 716;
  debounceMethod : USINT := TIME_UP_DOWN;
END_STRUCT;
END_TYPE

TYPE DFC_rbr_outK87OT : STRUCT
  DTC : UDINT := 16#046000;
  DFCid : UINT := 717;
  debounceMethod : USINT := TIME_UP_DOWN;
END_STRUCT;
END_TYPE

TYPE DFC_rbr_outK73SCB : STRUCT
  DTC : UDINT := 16#044100;
  DFCid : UINT := 686;
  debounceMethod : USINT := TIME_UP_DOWN;
END_STRUCT;
END_TYPE

TYPE DFC_rbr_outK73SCG : STRUCT
  DTC : UDINT := 16#044200;
  DFCid : UINT := 687;
  debounceMethod : USINT := TIME_UP_DOWN;
END_STRUCT;
END_TYPE

TYPE DFC_rbr_outK73OL : STRUCT
  DTC : UDINT := 16#043E00;
  DFCid : UINT := 683;
  debounceMethod : USINT := TIME_UP_DOWN;
END_STRUCT;
END_TYPE

TYPE DFC_rbr_outK73OT : STRUCT
  DTC : UDINT := 16#044000;
  DFCid : UINT := 685;
  debounceMethod : USINT := TIME_UP_DOWN;
END_STRUCT;
END_TYPE

TYPE DFC_rbr_outK73OC : STRUCT
  DTC : UDINT := 16#043D00;
  DFCid : UINT := 1053;
  debounceMethod : USINT := NO_DEBOUNCE;
END_STRUCT;
END_TYPE

TYPE DFC_rbr_outK73OR : STRUCT
  DTC : UDINT := 16#043F00;
  DFCid : UINT := 684;
  debounceMethod : USINT := TIME_UP_DOWN;
END_STRUCT;
END_TYPE

TYPE DFC_rbr_outK08SCB : STRUCT
  DTC : UDINT := 16#040B00;
  DFCid : UINT := 633;
  debounceMethod : USINT := TIME_UP_DOWN;
END_STRUCT;
END_TYPE

TYPE DFC_rbr_outK08SCG : STRUCT
  DTC : UDINT := 16#040C00;
  DFCid : UINT := 634;
  debounceMethod : USINT := TIME_UP_DOWN;
END_STRUCT;
END_TYPE

TYPE DFC_rbr_outK08OL : STRUCT
  DTC : UDINT := 16#040800;
  DFCid : UINT := 630;
  debounceMethod : USINT := TIME_UP_DOWN;
END_STRUCT;
END_TYPE

TYPE DFC_rbr_outK08OT : STRUCT
  DTC : UDINT := 16#040A00;
  DFCid : UINT := 632;
  debounceMethod : USINT := TIME_UP_DOWN;
END_STRUCT;
END_TYPE

TYPE DFC_rbr_outK08OC : STRUCT
  DTC : UDINT := 16#040700;
  DFCid : UINT := 1033;
  debounceMethod : USINT := NO_DEBOUNCE;
END_STRUCT;
END_TYPE

TYPE DFC_rbr_outK08OR : STRUCT
  DTC : UDINT := 16#040900;
  DFCid : UINT := 631;
  debounceMethod : USINT := TIME_UP_DOWN;
END_STRUCT;
END_TYPE

TYPE DFC_rbr_outK07SCB : STRUCT
  DTC : UDINT := 16#040500;
  DFCid : UINT := 628;
  debounceMethod : USINT := TIME_UP_DOWN;
END_STRUCT;
END_TYPE

TYPE DFC_rbr_outK07SCG : STRUCT
  DTC : UDINT := 16#040600;
  DFCid : UINT := 629;
  debounceMethod : USINT := TIME_UP_DOWN;
END_STRUCT;
END_TYPE

TYPE DFC_rbr_outK07OL : STRUCT
  DTC : UDINT := 16#040200;
  DFCid : UINT := 625;
  debounceMethod : USINT := TIME_UP_DOWN;
END_STRUCT;
END_TYPE

TYPE DFC_rbr_outK07OT : STRUCT
  DTC : UDINT := 16#040400;
  DFCid : UINT := 627;
  debounceMethod : USINT := TIME_UP_DOWN;
END_STRUCT;
END_TYPE

TYPE DFC_rbr_outK07OC : STRUCT
  DTC : UDINT := 16#040100;
  DFCid : UINT := 1031;
  debounceMethod : USINT := NO_DEBOUNCE;
END_STRUCT;
END_TYPE

TYPE DFC_rbr_outK07OR : STRUCT
  DTC : UDINT := 16#040300;
  DFCid : UINT := 626;
  debounceMethod : USINT := TIME_UP_DOWN;
END_STRUCT;
END_TYPE

TYPE DFC_rbr_outK29SCB : STRUCT
  DTC : UDINT := 16#043300;
  DFCid : UINT := 674;
  debounceMethod : USINT := TIME_UP_DOWN;
END_STRUCT;
END_TYPE

TYPE DFC_rbr_outK29SCG : STRUCT
  DTC : UDINT := 16#043400;
  DFCid : UINT := 675;
  debounceMethod : USINT := TIME_UP_DOWN;
END_STRUCT;
END_TYPE

TYPE DFC_rbr_outK29OL : STRUCT
  DTC : UDINT := 16#043000;
  DFCid : UINT := 671;
  debounceMethod : USINT := TIME_UP_DOWN;
END_STRUCT;
END_TYPE

TYPE DFC_rbr_outK29OT : STRUCT
  DTC : UDINT := 16#043200;
  DFCid : UINT := 673;
  debounceMethod : USINT := TIME_UP_DOWN;
END_STRUCT;
END_TYPE

TYPE DFC_rbr_outK29OC : STRUCT
  DTC : UDINT := 16#042F00;
  DFCid : UINT := 1049;
  debounceMethod : USINT := NO_DEBOUNCE;
END_STRUCT;
END_TYPE

TYPE DFC_rbr_outK29OR : STRUCT
  DTC : UDINT := 16#043100;
  DFCid : UINT := 672;
  debounceMethod : USINT := TIME_UP_DOWN;
END_STRUCT;
END_TYPE

TYPE DFC_rbr_outK09SCB : STRUCT
  DTC : UDINT := 16#041100;
  DFCid : UINT := 638;
  debounceMethod : USINT := TIME_UP_DOWN;
END_STRUCT;
END_TYPE

TYPE DFC_rbr_outK09SCG : STRUCT
  DTC : UDINT := 16#041200;
  DFCid : UINT := 639;
  debounceMethod : USINT := TIME_UP_DOWN;
END_STRUCT;
END_TYPE

TYPE DFC_rbr_outK09OL : STRUCT
  DTC : UDINT := 16#040E00;
  DFCid : UINT := 635;
  debounceMethod : USINT := TIME_UP_DOWN;
END_STRUCT;
END_TYPE

TYPE DFC_rbr_outK09OT : STRUCT
  DTC : UDINT := 16#041000;
  DFCid : UINT := 637;
  debounceMethod : USINT := TIME_UP_DOWN;
END_STRUCT;
END_TYPE

TYPE DFC_rbr_outK09OC : STRUCT
  DTC : UDINT := 16#040D00;
  DFCid : UINT := 1035;
  debounceMethod : USINT := NO_DEBOUNCE;
END_STRUCT;
END_TYPE

TYPE DFC_rbr_outK09OR : STRUCT
  DTC : UDINT := 16#040F00;
  DFCid : UINT := 636;
  debounceMethod : USINT := TIME_UP_DOWN;
END_STRUCT;
END_TYPE

TYPE DFC_rbr_outK51SCB : STRUCT
  DTC : UDINT := 16#043800;
  DFCid : UINT := 678;
  debounceMethod : USINT := TIME_UP_DOWN;
END_STRUCT;
END_TYPE

TYPE DFC_rbr_outK51SCG : STRUCT
  DTC : UDINT := 16#043900;
  DFCid : UINT := 679;
  debounceMethod : USINT := TIME_UP_DOWN;
END_STRUCT;
END_TYPE

TYPE DFC_rbr_outK51OL : STRUCT
  DTC : UDINT := 16#043600;
  DFCid : UINT := 676;
  debounceMethod : USINT := TIME_UP_DOWN;
END_STRUCT;
END_TYPE

TYPE DFC_rbr_outK51OT : STRUCT
  DTC : UDINT := 16#043700;
  DFCid : UINT := 677;
  debounceMethod : USINT := TIME_UP_DOWN;
END_STRUCT;
END_TYPE

TYPE DFC_rbr_outK51OC : STRUCT
  DTC : UDINT := 16#043500;
  DFCid : UINT := 1051;
  debounceMethod : USINT := NO_DEBOUNCE;
END_STRUCT;
END_TYPE

TYPE DFC_rbr_outK14SCB : STRUCT
  DTC : UDINT := 16#042000;
  DFCid : UINT := 651;
  debounceMethod : USINT := TIME_UP_DOWN;
END_STRUCT;
END_TYPE

TYPE DFC_rbr_outK14SCG : STRUCT
  DTC : UDINT := 16#042100;
  DFCid : UINT := 652;
  debounceMethod : USINT := TIME_UP_DOWN;
END_STRUCT;
END_TYPE

TYPE DFC_rbr_outK14OL : STRUCT
  DTC : UDINT := 16#041E00;
  DFCid : UINT := 648;
  debounceMethod : USINT := TIME_UP_DOWN;
END_STRUCT;
END_TYPE

TYPE DFC_rbr_outK14OT : STRUCT
  DTC : UDINT := 16#041F00;
  DFCid : UINT := 650;
  debounceMethod : USINT := TIME_UP_DOWN;
END_STRUCT;
END_TYPE

TYPE DFC_rbr_outK14OC : STRUCT
  DTC : UDINT := 16#041D00;
  DFCid : UINT := 1041;
  debounceMethod : USINT := NO_DEBOUNCE;
END_STRUCT;
END_TYPE

TYPE DFC_rbr_outK80SCB : STRUCT
  DTC : UDINT := 16#044500;
  DFCid : UINT := 690;
  debounceMethod : USINT := TIME_UP_DOWN;
END_STRUCT;
END_TYPE

TYPE DFC_rbr_outK80SCG : STRUCT
  DTC : UDINT := 16#044600;
  DFCid : UINT := 691;
  debounceMethod : USINT := TIME_UP_DOWN;
END_STRUCT;
END_TYPE

TYPE DFC_rbr_outK80OL : STRUCT
  DTC : UDINT := 16#044300;
  DFCid : UINT := 688;
  debounceMethod : USINT := TIME_UP_DOWN;
END_STRUCT;
END_TYPE

TYPE DFC_rbr_outK80OT : STRUCT
  DTC : UDINT := 16#044400;
  DFCid : UINT := 689;
  debounceMethod : USINT := TIME_UP_DOWN;
END_STRUCT;
END_TYPE

TYPE DFC_rbr_outK81SCB : STRUCT
  DTC : UDINT := 16#044900;
  DFCid : UINT := 694;
  debounceMethod : USINT := TIME_UP_DOWN;
END_STRUCT;
END_TYPE

TYPE DFC_rbr_outK81SCG : STRUCT
  DTC : UDINT := 16#044A00;
  DFCid : UINT := 695;
  debounceMethod : USINT := TIME_UP_DOWN;
END_STRUCT;
END_TYPE

TYPE DFC_rbr_outK81OL : STRUCT
  DTC : UDINT := 16#044700;
  DFCid : UINT := 692;
  debounceMethod : USINT := TIME_UP_DOWN;
END_STRUCT;
END_TYPE

TYPE DFC_rbr_outK81OT : STRUCT
  DTC : UDINT := 16#044800;
  DFCid : UINT := 693;
  debounceMethod : USINT := TIME_UP_DOWN;
END_STRUCT;
END_TYPE

TYPE DFC_rbr_outK82SCB : STRUCT
  DTC : UDINT := 16#044D00;
  DFCid : UINT := 698;
  debounceMethod : USINT := TIME_UP_DOWN;
END_STRUCT;
END_TYPE

TYPE DFC_rbr_outK82SCG : STRUCT
  DTC : UDINT := 16#044E00;
  DFCid : UINT := 699;
  debounceMethod : USINT := TIME_UP_DOWN;
END_STRUCT;
END_TYPE

TYPE DFC_rbr_outK82OL : STRUCT
  DTC : UDINT := 16#044B00;
  DFCid : UINT := 696;
  debounceMethod : USINT := TIME_UP_DOWN;
END_STRUCT;
END_TYPE

TYPE DFC_rbr_outK82OT : STRUCT
  DTC : UDINT := 16#044C00;
  DFCid : UINT := 697;
  debounceMethod : USINT := TIME_UP_DOWN;
END_STRUCT;
END_TYPE

TYPE DFC_rbr_outK83SCB : STRUCT
  DTC : UDINT := 16#045100;
  DFCid : UINT := 702;
  debounceMethod : USINT := TIME_UP_DOWN;
END_STRUCT;
END_TYPE

TYPE DFC_rbr_outK83SCG : STRUCT
  DTC : UDINT := 16#045200;
  DFCid : UINT := 703;
  debounceMethod : USINT := TIME_UP_DOWN;
END_STRUCT;
END_TYPE

TYPE DFC_rbr_outK83OL : STRUCT
  DTC : UDINT := 16#044F00;
  DFCid : UINT := 700;
  debounceMethod : USINT := TIME_UP_DOWN;
END_STRUCT;
END_TYPE

TYPE DFC_rbr_outK83OT : STRUCT
  DTC : UDINT := 16#045000;
  DFCid : UINT := 701;
  debounceMethod : USINT := TIME_UP_DOWN;
END_STRUCT;
END_TYPE

TYPE DFC_rbr_outK25SCB : STRUCT
  DTC : UDINT := 16#042D00;
  DFCid : UINT := 669;
  debounceMethod : USINT := TIME_UP_DOWN;
END_STRUCT;
END_TYPE

TYPE DFC_rbr_outK25SCG : STRUCT
  DTC : UDINT := 16#042E00;
  DFCid : UINT := 670;
  debounceMethod : USINT := TIME_UP_DOWN;
END_STRUCT;
END_TYPE

TYPE DFC_rbr_outK25OR : STRUCT
  DTC : UDINT := 16#042C00;
  DFCid : UINT := 668;
  debounceMethod : USINT := TIME_UP_DOWN;
END_STRUCT;
END_TYPE

TYPE DFC_rbr_outK62SCB : STRUCT
  DTC : UDINT := 16#043B00;
  DFCid : UINT := 681;
  debounceMethod : USINT := TIME_UP_DOWN;
END_STRUCT;
END_TYPE

